        | 	pivot_pose = pose_trans(p_center, hinge_offset)
        | 	pose_rel = pose_trans(pose_inv(pivot_pose), p_center)
        | 	angle_mid = (angle/2.0)*3.1416/180
        | 	angle_end = angle*3.1416/180
        | 	tilt_mid = p[0,0,0, -angle_mid, 0, 0]
        | 	tilt_end = p[0,0,0, -angle_end, 0, 0]
        | 	pose_rel_mid = pose_trans(tilt_mid, pose_rel)
        | 	pose_rel_end = pose_trans(tilt_end, pose_rel)
        | 	via_pose = pose_trans(pivot_pose, pose_rel_mid)
        | 	end_pose = pose_trans(pivot_pose, pose_rel_end)
        | 	movec(via_pose, end_pose, a=0.05, v=0.01, r=0.001)
        | 	p_center = get_actual_tcp_pose()
        | end
        | 
        | def deg2rad(d):
        | 	return d*3.141592/180
        | end
        | 
        | def map_tilt_to_ry_deg(container_deg):
        | 
        | 	if (Flowability == "Easy" or Flowability == "Medium"):
        | 		if ( level>=10.0):
        | 			ry_min = 10.0
        | 			ry_max = 75.0
        | 		elif (level<10.00 and level >1.00):
        | 			ry_min = 16.0
        | 			ry_max = 65.0
        | 		else:
        | 			ry_min=17.0
        | 			ry_max=75.0
        | 		end
        | 	else:
        | 		if ( level>=10.0):
        | 			ry_min = 0.0
        | 			ry_max = 65.0
        | 		elif (level<10.00 and level >1.00):
        | 			ry_min = 10.0
        | 			ry_max = 45.0
        | 		else:
        | 			ry_min=0.0
        | 			ry_max=50.0
        | 		end
        | 
        | 	end
        | 
        | 	local span_count = angle_max -angle_min
        | 	local span_ry = ry_max - ry_min
        | 
        | 	local t = (container_deg -angle_min)/span_count
        | 	local ry_deg = ry_max - t*span_ry
        | 
        | 	return clamp(ry_deg, ry_min, ry_max)
        | 
        | end
        | 
        | def caluclate_corrections(level):
        | 	z_high = 0.01
        | 	z_low = -0.08
        | 	y_high = -0.01
        | 	y_low = -0.015
        | 
        | 	scale = (level - 10.0) / (100.0-10.0)
        | 
        | 	global correction_z = z_low + scale*(z_high - z_low)
        | 	global correction_y = y_low + scale*(y_high -y_low)
        | 
        | end
        | 
        | def scoop_powder(p_center):
        | 	#lift_offset = p[0, 0, 0.05, 0, 0, 0]
        | 	vibration_voltage = 0.4
        | 	vibration_time = 3.0
        | 	diameter = 0.07
        | 	global scoop_radius_default = 0.0
        | 	#p_center = center_pose_t
        | 
        | 
        | 	if (level >=70.00):
        | 		approach_offset = p[0.008,0,0.22,0,0,0]
        | 		lift_offset = p[0, 0, 0.05, 0, 0, 0]
        | 		caluclate_corrections(level)
        | 	elif (level >=10.00 and level <70):
        | 		approach_offset = p[0.008,0,0.22,0,0,0]
        | 		lift_offset = p[0, 0, 0.15, 0, 0, 0]
        | 		caluclate_corrections(level)
        | 	elif (level<10.00 and level >= 1.00):
        | 		approach_offset = p[0.01,0,0.22,0,0,0]
        | 		correction_z = -0.08
        | 		correction_y = -0.01
        | 		lift_offset = p[0, 0, 0.14, 0, 0, 0]
        | 	else:
        | 		approach_offset = p[0.008,0,0.22,0,0,0]
        | 		correction_z = -0.08
        | 		correction_y = -0.01
        | 		lift_offset = p[0, 0, 0.14, 0, 0, 0]
        |  	end
        | 
        | 	if (spatula == "spatula_L"):
        | 		global spatula_depth = 0.015
        | 	elif (spatula == "spatula_M"):
        | 		global spatula_depth = 0.01
        | 	elif (spatula == "spatula_S"):
        | 		global spatula_depth = 0.008
        | 	elif (spatula == "spatula_flat_M"):
        | 		global spatula_depth = 0.001
        | 	elif (spatula == "spatula_flat_S"):
        | 		global spatula_depth = 0.005
        | 	end
        | 
        | 	scoop_radius_default = diameter/2 - spatula_depth
        | 	scoop_entry_pose = pose_trans(p_center, approach_offset)
        | 	movel(scoop_entry_pose, a=0.1, v=0.25)
        | 
        | 	scoop_start_rel = p[scoop_radius_default, 0, scoop_depth, 0, 0, 0]
        | 
        | 	rot_mid = p[0, 0, 0, 0, 0, 0.785]
        | 	rot_end = p[0, 0, 0, 0, 0, 1.5708]
        | 
        | 	scoop_via_rel = pose_trans(rot_mid, scoop_start_rel)
        | 	scoop_end_rel = pose_trans(rot_end, scoop_start_rel)
        | 
        | 	scoop_start_pose = pose_trans(p_center, scoop_start_rel)
        | 	scoop_via_pose = pose_trans(p_center, scoop_via_rel)
        | 	scoop_end_pose = pose_trans(p_center, scoop_end_rel)
        | 
        | 	movel(scoop_start_pose, a=0.5, v=0.3)
        | 	#movel(p_center, a=0.5, v=1.0)
        | 	#sleep(5.0)
        | 
        | 	if (level<90.0):
        | 		Rotate()
        | 	end
        | 
        | 	#movec(scoop_via_pose, scoop_end_pose, a=0.03, v=0.05)
        | 	movec(scoop_via_pose, scoop_end_pose, a=0.03, v=0.02)
        | 	#movel(pose_trans(get_actual_tcp_pose(), p[0,0,0,0,0,deg2rad(90.0)]), a=0.03, v=0.05)
        | 	sleep(1.0)
        | 	local ry_deg = map_tilt_to_ry_deg(angle_deg)
        | 	local ry = deg2rad(ry_deg)
        | 	local end_rel = pose_trans(pose_inv(p_center), scoop_end_pose)
        | 	local end_rel_tilted = pose_trans(end_rel, p[0, 0, 0, 0, ry, 0])
        | 	global tilted_pose_in_base = pose_trans(p_center, p[0,correction_y,correction_z,end_rel_tilted[3],end_rel_tilted[4], end_rel_tilted[5]])
        | 	global tilted_pose_in_base = pose_trans(tilted_pose_in_base, p[0, 0, spatula_len, 0, 0, 0])
        | 
        | 	if (Flowability == "Hard"):
        | 		tilt_send((angle_deg+5))
        | 	end
        | 	movel(tilted_pose_in_base, a=0.03, v=0.1)
        | 
        | 	if (Flowability == "Hard"):
        | 		tilt_send((angle_deg-5))
        | 	end
        | 
        | 	if (spatula=="spatula_flat_S" or spatula=="spatula_S"):
        | 		vibration_3()
        | 	else:
        | 		set_analog_out(0, vibration_voltage)
        | 	end
        | 	if (Flowability == "Easy"):
        | 		local n=1.4
        | 	else:
        | 		local n=1.5
        | 	end
        | 	local ry_level = deg2rad(ry_deg/n)
        | 	local end_rel_tilted_level = pose_trans(end_rel, p[0, 0, 0, 0, ry_level, 0])
        | 	local level_tilted_pose_in_base = pose_trans(p_center, p[0,correction_y,correction_z,end_rel_tilted_level[3],end_rel_tilted_level[4], end_rel_tilted_level[5]])
        | 	local level_tilted_pose_in_base = pose_trans(level_tilted_pose_in_base, p[0, 0, spatula_len, 0, 0, 0])
        | 
        | 	movel(level_tilted_pose_in_base, a=0.03, v=0.1)
        | 	#if (level>70.0):
        | 		#sleep(1.0)
        | 	#end
        | 	sleep(1.0)
        | 	#sleep(vibration_time)
        | 
        | 	movel(tilted_pose_in_base, a=0.03, v=0.1)
        | 	set_analog_out(0, 0.0)
        | 
        | 	tilt_pose_rel = pose_trans(pose_inv(p_center), tilted_pose_in_base)
        | 
        | 	lifted_pose_rel = pose_trans(lift_offset, tilt_pose_rel)
        | 
        | 	global lifted_pose = pose_trans(p_center, lifted_pose_rel)
        | 	movel(lifted_pose, a=0.03, v=0.1)
        | 	CCW_Rotate()
        | end
        | 
        | 
        | def center_pose():
        | 	trans_rel = p[0.0, 0.05, 0.0, 0, 0, 0]
        | 
        | 	p_translated = pose_trans(place_pose, trans_rel)
        | 	cx = p_translated[0]
        | 	cy = p_translated[1]
        | 	cz = p_translated[2]
        | 
        | 	global p_center_vertical = p[cx,cy,cz, 0, 0, 4.09]
        | 
        | 	#movej(p_center_vertical, a =0.3, v =0.3)
        | 	#sleep(3.0)
        | 	return p_center_vertical
        | end
        | 
        | def updated_center_pose(p_center_vertical, angle_deg):
        | 	hinge_pose = pose_trans(p_center_vertical, p[0,0,-0.2,0,0,0])
        | 	local_rel = pose_trans(pose_inv(hinge_pose), p_center_vertical)
        | 
        | 	rot_tilt = p[0,0,0, -deg2rad(angle_deg),0,0]
        | 	local_rel_tilted = pose_trans(rot_tilt, local_rel)
        | 
        | 	global p_center = pose_trans(hinge_pose, local_rel_tilted)
        | 	return p_center
        | end
        | 
        | def tilt_send(angle):
        | 	socket_open("192.168.12.101", 80)
        | 	angle = 92.0 - angle
        | 	socket_send_string("Tilt,"+to_str(angle)+",0")
        | 	sync()
        | 	sleep(0.5)
        | 	socket_close()
        | end
        | 
        | def Motors_off():
        | 	socket_open("192.168.12.101", 80)
        | 	socket_send_string("Off,0,0")
        | 	sync()
        | 	sleep(0.5)
        | 	socket_close()
        | end
        | 
        | def Rotate():
        | 	socket_open("192.168.12.101", 80)
        | 	socket_send_string("FullRotation, 1, 2000")
        | 	sync()
        | 	sleep(0.5)
        | 	socket_close()
        | end
        | 
        | 
        | def CCW_Rotate():
        | 	socket_open("192.168.12.101", 80)
        | 	socket_send_string("FullRotation, -1, 2000")
        | 	sync()
        | 	sleep(0.5)
        | 	socket_close()
        | end
        | def tilt_to_home():
        | 	socket_open("192.168.12.101", 80)
        | 	socket_send_string("Home,0,0")
        | 	sync()
        | 	sleep(0.5)
        | 	socket_close()
        | end
    Script file /programs/04 Scripts/Weight_scale_socket.script
      | def get_weight():
      | 	socket_open("192.168.12.111", 3002)
      | 	sleep(0.2)
      | 	textmsg("socket opened successfully!")
      | 	socket_send_string("GET_WEIGHT")
      | 	sync()
      | 	sleep(0.5)
      | 	receiveFromServ = socket_read_ascii_float(6)
      | 	while (receiveFromServ[0] <1):
      | 		sleep(0.5)
      | 		receiveFromServ = socket_read_ascii_float(1)
      | 		textmsg("retrying read:", receiveFromServ)
      | 	end
      | 	textmsg("Received weight:", receiveFromServ[1])
      | 	socket_close()
      | 	sleep(0.2)
      | 	return receiveFromServ[1]
      | end
      | 
      | def tare_scale():
      | 	socket_open("192.168.12.111", 3002)
      | 	socket_send_string("TARE")
      | 	sleep(0.5)
      | 	socket_close()
      | end
      | 
      | def zero_scale():
      | 	socket_open("192.168.12.111", 3002)
      | 	socket_send_string("ZERO")
      | 	sleep(0.5)
      | 	socket_close()
      | end
      | 
      | def log_weight():
      | 	socket_open("192.168.12.111", 3002)
      | 	socket_send_string("LOG_WEIGHT")
      | 	sleep(0.5)
      | 	socket_close()
      | end
      | 
      | def send_target_info():
      | 	socket_open("192.168.12.111", 3002)
      | 	socket_send_string("SET_TARGET:" + to_str(target_weight))
      | 	sleep(0.2)
      | 	socket_close()
      | end
      | def send_powder_info():
      | 	socket_open("192.168.12.111", 3002)
      | 	socket_send_string("SET_POWDER:" + Pow_name)
      | 	sleep(0.2)
      | 	socket_close()
      | end
      | def send_spatula_info():
      | 	socket_open("192.168.12.111", 3002)
      | 	socket_send_string("SET_SPATULA:" + spatula)
      | 	sleep(0.2)
      | 	socket_close()
      | end
      | 
      | def send_level_info():
      | 	socket_open("192.168.12.111", 3002)
      | 	socket_send_string("SET_LEVEL:" + to_str(level))
      | 	sleep(0.2)
      | 	socket_close()
      | end
      | def Dosing_done():
      | 	socket_open("192.168.12.111", 3002)
      | 	socket_send_string("DOSING_DONE")
      | 	sleep(0.2)
      | 	socket_close()
      | end
      | 
      | def send_dosing_time(Dosed_time):
      | 	socket_open("192.168.12.111", 3002)
      | 	socket_send_string("DOSED_TIME:" + to_str(Dosed_time))
      | 	sleep(0.2)
      | 	socket_close()
      | end
    Script file /programs/04 Scripts/Calibration.script
      | # ------------------------------------------------------------
      | # Theoretical W_FULL from Cylinder Volume + Density
      | # (Eliminates manual W_FULL; keeps W_EMPTY + W_now for level)
      | # ------------------------------------------------------------
      | # -------------------------
      | # 1) Define container geometry (cylindrical inner dimensions)
      | # -------------------------
      | # Use mm for readability; we convert internally.
      | global D_INNER_MM   = 66.0     # inner diameter of container (mm)
      | global H_FILL_MM    = 125.0    # usable fill height up to "full" (mm)
      | 
      | # -------------------------
      | # 2) Define powder density
      | # -------------------------
      | # Density is directly set for now (as per your requirement).
      | # Use g/mL (common lab bulk density style).
      | #global RHO_G_PER_ML = 0.40     # example: 0.55 g/mL (replace per powder)
      | 
      | # ------------------------------------------------------------
      | # Spatula volumes (manufacturer specified)
      | # ------------------------------------------------------------
      | 
      | # Large spatula
      | global SPATULA_L_VOL_ML = 5.0        # 1 teaspoon = 5 mL
      | 
      | # Medium spatula
      | global SPATULA_M_VOL_ML = 1.25       # 1/4 teaspoon = 1.25 mL
      | 
      | # Small spatula
      | global SPATULA_S_VOL_ML = 0.15625    # 1/32 teaspoon = 0.15625 mL
      | 
      | global SPATULA_FLAT_M_VOL_ML  = 2.2
      | global SPATULA_FLAT_S_VOL_ML  = 1.2   #based on caluclations using rho = m/V
      | 
      | # -------------------------
      | # 4) Utility functions
      | # -------------------------
      | 
      | 
      | def cyl_volume_mL(d_mm, h_mm):
      |   # Converts mm -> m, computes cylinder volume in m^3, converts to mL
      |   # V = π * r^2 * h
      |   local d_m  = d_mm / 1000.0
      |   local h_m  = h_mm / 1000.0
      |   local r_m  = d_m / 2.0
      |   local v_m3 = 3.141592653589793 * r_m * r_m * h_m
      |   global v_mL = v_m3 * 1000000.0     # 1 m^3 = 1,000,000 mL
      |   return v_mL
      | end
      | 
      | def compute_W_full_theoretical():
      |   V_mL = cyl_volume_mL(D_INNER_MM, H_FILL_MM)
      |   local M_powder_g = density * V_mL
      |   global W_FULL = W_EMPTY + M_powder_g
      |   return W_FULL
      | end
      | 
      | 
      | # ------------------------------------------------------------
      | # Function: Theoretical scoop weight from volume
      | # ------------------------------------------------------------
      | def scoop_weight_from_volume(vol_mL, density):
      |   return vol_mL * density
      | end
      | 
      | # ------------------------------------------------------------
      | # Function: Get scoop weight based on spatula type
      | # ------------------------------------------------------------
      | def get_scoop_weight(spatula):
      |   local vol = 0.0
      | 
      |   if (spatula == "spatula_L"):
      |     vol = SPATULA_L_VOL_ML
      |   elif (spatula == "spatula_M"):
      |     vol = SPATULA_M_VOL_ML
      |   elif (spatula == "spatula_S"):
      |     vol = SPATULA_S_VOL_ML
      |   elif (spatula == "spatula_flat_M"):
      |     return SPATULA_FLAT_M_VOL_ML
      |   elif (spatula == "spatula_flat_S"):
      |     return SPATULA_FLAT_S_VOL_ML
      |   else:
      |     textmsg("Unknown spatula type")
      |     return 0.0
      |   end
      | 
      |   global target_g =  scoop_weight_from_volume(vol, density)
      |   return target_g
      | end
  Folder BeforeStarts [hidden by the author, left out]
  Folder powder dispensing variable init
    Start_thread := False
    vib_thread := False
    kp := 0.001
    ki := 0.00006
    kd := 0.015
    dt := 0.03
    Integral_error := 0
    current_error := 0
    previous_error := 0
    tilt_increment := 0
    tilt_angle := 0
    diff := 0
    current_pose := get_actual_tcp_pose()
    Relative_trans := p[0, 0, -0.035, 0, 0, 0]
    ContA_plc_offst := p[-0.00205, 0.02547, 0.03730, -0.03, -2.183, 6.165]
    PowA_50_offset := p[0.21808, -0.19943, 0.06584, 0, 0, 0]
    SuppressedNode
      Script: scooping_init()
    Script: tilt_init_reference()
    switch_spat_M := True
    switch_spat_S := True
    switch_spat_F_M := True
    switch_spat_F_S := True
    last_scale := 0
    W_EMPTY := 51.3
    w_dosed_total := 0
Robot Program (runOnlyOnce=false)
  Folder MAIN
    Script: command_manager(external_control="uGO", cond_suspend=(ITM_Manipulated and AMR_AtTarget and AMR_Charging and AMR_Battery<40), cond_unsuspend=(AMR_Battery≟60))
    Script: log_state(STATE_Info)
    Switch expression=STATE
      Case (caseValue=1)
        Folder Stopping
          STATE_Info := "Stopping"
          Script: end_freedrive_mode()
          Set NoAction tcp=TCP
          PSE_T := get_tool_free_pose(dir=[0,0,0.150], move_in_base_frame=True)
          If is_reachable(Base, [PSE_T])
            MoveL speed 150 mm/s, acceleration 1200 mm/s^2 (useActiveTCP=true optimoveEnabled=false optiMoveSpeed=0.3 optiMoveAcceleration=0.09) feature=Base
              Waypoint Variable (Variable): variable=PSE_T
          Script: do_transition(keep_rxry=OBJ_Picked, r=0)
          SuppressedNode
            Folder Decapper
              Set DigitalOutput pin=digital_out[4]; digitalValue=0
              Set DigitalOutput pin=BarcodeTrigger; digitalValue=0
              Set DigitalOutput pin=digital_out[3]; digitalValue=0
              Set DigitalOutput pin=digital_out[2]; digitalValue=0
              Set DigitalOutput pin=digital_out[5]; digitalValue=0
          SuppressedNode
            Folder Centrifuge [hidden by the author, left out]
          Call Sub_AMR_MiR_V3
          If stopping() and AMR_Done
            STATE := 2
            Script: ugo_update_outputs()
      Case (caseValue=2)
        Folder Stopped
          STATE_Info := "Stopped"
          Call Sub_AMR_MiR_V3
          If CMD_Reset  or PB_Start
            STATE := 3
            Script: ugo_update_outputs()
      Case (caseValue=3)
        Folder  Resetting [hidden by the author, left out]
      Case (caseValue=4)
        Folder Idle [hidden by the author, left out]
      Case (caseValue=5)
        Folder Starting
          STATE_Info := "Starting"
          'ADD COMMANDS WHAT TO START WITH'
          Call Sub_AMR_MiR_V3
          Folder get ugo data
            Folder Assign Tasks
              Script: TASK.ID = ugo_get_task()
              If TASK.ID≟1
                Task_info := "Charge"
                Folder Parameters
                  AMR_PosTarget := 1
              ElseIf TASK.ID≟9
                'Pick Sarstedt Rack from Variable source'
                Task_info := "Navigate to Target"
                Folder Parameters
                  AMR_PosTarget := UGO.read_input("00","ITM_ID")
              ElseIf TASK.ID≟49
                Task_info := "Pick Containers"
                Folder Parameters
                  ITM_ID := 1
                  OBJ_Type := 6
                  JIG := 15
                  AMR_PosTarget := 3
              ElseIf TASK.ID≟50
                Task_info := "Decap Containers"
                Folder Parameters
                  ITM_ID := 1
                  OBJ_Type := 6
                  JIG := 16
                  AMR_PosTarget := 5
              ElseIf TASK.ID≟51
                Task_info := "Detect Spatula and transfer powder"
                Folder Parameters
                  ITM_ID := 1
                  target_weight := (UGO.read_input("00","Target_weight"))/1000
                  OBJ_Type := 8
                  JIG := 16
                  AMR_PosTarget := 5
              ElseIf TASK.ID≟52
                Task_info := "Pick Powder"
                Folder Parameters
                  ITM_ID := 1
                  OBJ_Type := 6
                  JIG := 15
                  AMR_PosTarget := 3
              ElseIf TASK.ID≟53
                Task_info := "Decap Powder"
                Folder Parameters
                  ITM_ID := 1
                  OBJ_Type := 6
                  JIG := 1
                  AMR_PosTarget := 5
              ElseIf TASK.ID≟54
                Task_info := "Empty and swap Powder container"
                SuppressedNode
                  Folder Parameters
                    ITM_ID := 1
                    target_weight := (UGO.read_input("00","Target_weight"))/1000
                    W_now := (UGO.read_input("00","Container_weight"))/1000
                    Pow_name := (UGO.read_input("00","Powder_name"))
                    OBJ_Type := 6
                    JIG := 17
                    AMR_PosTarget := 5
                Folder Parameters
                  ITM_ID := 1
                  SuppressedNode
                    target_weight := (UGO.read_input("00","target_weight"))/1000
                  W_now := (UGO.read_input("00","Container_weight"))/1000
                  Pow_name := (UGO.read_input("00","Powder_name"))
                  Script: scooping_init()
                  target_weight := W_now-W_EMPTY-(0.002*W_FULL)
                  OBJ_Type := 6
                  JIG := 17
                  AMR_PosTarget := 5
              ElseIf TASK.ID≟55
                Task_info := "Place Powder"
                Folder Parameters
                  ITM_ID := 1
                  OBJ_Type := 6
                  JIG := 21
                  AMR_PosTarget := 5
              ElseIf TASK.ID≟56
                Task_info := "Dose Powder"
                Folder Parameters
                  ITM_ID := 1
                  target_weight := (UGO.read_input("00","Target_weight"))/1000
                  W_now := (UGO.read_input("00","Container_weight"))/1000
                  SuppressedNode
                    W_now := 135
                  Pow_name := (UGO.read_input("00","Powder_name"))
                  OBJ_Type := 6
                  JIG := 17
                  AMR_PosTarget := 5
              ElseIf TASK.ID≟57
                Task_info := "Recipe Powder dosing"
                Folder Parameters
                  ITM_ID := 1
                  Pow_A := (UGO.read_input("00","PowderA"))
                  Pow_B := (UGO.read_input("00","PowderB"))
                  Pow_C := (UGO.read_input("00","PowderC"))
                  Total_weight := (UGO.read_input("00","Total_weight"))/1000
                  Pow_A_percent := (UGO.read_input("00","PowderA_percentage"))/100
                  Pow_B_percent := (UGO.read_input("00","PowderB_percentage"))/100
                  Pow_C_percent := (UGO.read_input("00","PowderC_percentage"))/100
                  OBJ_Type := 6
                  JIG := 17
                  AMR_PosTarget := 5
              ElseIf TASK.ID≟58
                Task_info := "Pick Powder containers"
                Folder Parameters
                  ITM_ID := 1
                  OBJ_Type := 6
                  JIG := 15
                  AMR_PosTarget := 3
              ElseIf TASK.ID≟59
                Task_info := "Calibration for new powder"
                Folder Parameters
                  ITM_ID := 1
                  Pow_name := (UGO.read_input("00","Pow_name"))
                  W_now := (UGO.read_input("00","Container_weight"))/1000
                  density := (UGO.read_input("00", "Density"))
                  Flowability := (UGO.read_input("00", "Flowability"))
                  spatula := (UGO.read_input("00","Spatula"))
                  OBJ_Type := 6
                  JIG := 17
                  AMR_PosTarget := 5
              Else 
                Script: set_error(ERROR_WRONG_ORDER)
          Folder test ugo
            Wait Sleep waitTime=0.2
            Script: ugo_update_outputs()
          If starting() and AMR_Done
            Script: log_message(Task_info, "New Task: ")
            Script: log_message(to_str(TASK.ID), "Task_ID: ")
            Script: do_transition(keep_rxry=OBJ_Picked)
            STATE := 6
            Script: ugo_update_outputs()
      Case (caseValue=6)
        Folder Execute
          STATE_Info := "Execute"
          If not CMD_Hold and not CMD_Suspend (checkContinuously=true)
            Switch expression=PROCESS_Step
              Case (caseValue=0)
                PROCESS_Info := "process control"
                Script: log_process(PROCESS_Info)
                Folder process control [hidden by the author, left out]
              Case (caseValue=1)
                Folder navigate
                  'MOVING THE uML'
                  PROCESS_Info := "move to target"
                  Script: log_process(PROCESS_Info)
                  If TASK.ID≟1
                    Action := 51
                  Else 
                    Action := 52
                  Call Sub_AMR_MiR_V3
                  If AMR_Done
                    PROCESS_Step := 0
              Case (caseValue=2)
                Folder prepare
                  'THINGS THAT HAVE TO BE DONE ONCE IN A SEQUENCE,WORKFLOW'
                  PROCESS_Info := "prepare for work"
                  Script: log_process(PROCESS_Info)
                  If TASK.WORK.ITM_ID_Src>1
                    ITM_ID := TASK.WORK.ITM_ID_Src
                  ElseIf TASK.WORK.ITM_ID_Tgt>1
                    ITM_ID := TASK.WORK.ITM_ID_Tgt
                  If not ARM_Referenced and (ITM_ID≠0)
                    STP := 1
                  ElseIf ARM_Referenced or (ITM_ID≟0)
                    STP := 2
                  Switch expression=STP
                    Case (caseValue=1)
                      Folder reference
                        STP_Info := "reference at target position"
                        Script: log_step(STP_Info)
                        If ITM_ID≟1
                          CAM_Done := True
                        Else 
                          Action := 131
                          Call Sub_Vision_V18
                          SuppressedNode
                            CAM_Done := True
                        If CAM_Done and  not ERROR.FLAG
                          Script: log_step("ARM referenced")
                          ARM_Referenced := True
                    Case (caseValue=2)
                      Folder manipulate [hidden by the author, left out]
                  ITM_Prepared := (ITM_Manipulated or  not found_in_list(ITM_ID, ITM_ID_List)) and (ARM_Referenced or ITM_ID≟0) and  not WRK_Done
                  STP := 0
                  STP_Info := ""
                  PROCESS_Step := 0
              Case (caseValue=3)
                Folder work
                  'ADD EVERY MACHINE, OBJECT, STATION TO WORK ON'
                  Switch expression=ITM_ID
                    Case (caseValue=1)
                      Folder uLM
                        If TASK.ID≟12
                          Folder fill racks
                            Action := 151
                            Call Sub_Vision_V18
                            If not ERROR.FLAG
                              Folder Actions for the task
                                Action := 1
                                JIG := 2
                                JIG_Slot := CAM_Result[0]
                                OBJ_Nbr := CAM_Result[0]
                                OBJ_Type := 2
                                Call Sub_Action_V4
                                If OBJ_Picked
                                  Script: CAM_Result.remove(0)
                                  PRC_TubCounter := PRC_TubCounter+1
                                  If PRC_TubCounter%4≟0
                                    JIG_Slot := 4
                                  Else 
                                    JIG_Slot := PRC_TubCounter%4
                                  OBJ_Nbr := ceil(PRC_TubCounter/4)
                                  Action := 2
                                  JIG := 4
                                  Call Sub_Action_V4
                                  Action := 151
                                  Call Sub_Vision_V18
                            If (CAM_Captures≥CAM_PRM_Retries) or (PRC_TubCounter≥32)
                              PROCESS_Step := 0
                              WRK_Done := True
                        ElseIf TASK.ID≟49
                          Folder Pick Powder container
                            Action := 131
                            Call Sub_Vision_V18
                            Action := 35
                            Call Sub_Action_V4
                            PROCESS_Step := 0
                            WRK_Done := True
                        ElseIf TASK.ID≟50
                          Folder Decap containers
                            Action := 36
                            Call Sub_Action_V4
                            PROCESS_Step := 0
                            WRK_Done := True
                        ElseIf TASK.ID≟51
                          Folder Detect Spatula and transfer powder
                            Action := 131
                            Call Sub_Vision_V18
                            Action := 37
                            Call Sub_Action_V4
                            PROCESS_Step := 0
                            WRK_Done := True
                        ElseIf TASK.ID≟52
                          Folder Pick Powder container
                            Action := 131
                            Call Sub_Vision_V18
                            Action := 39
                            Call Sub_Action_V4
                            PROCESS_Step := 0
                            WRK_Done := True
                        ElseIf TASK.ID≟53
                          Folder Decap containerA
                            Action := 40
                            Call Sub_Action_V4
                            PROCESS_Step := 0
                            WRK_Done := True
                        ElseIf TASK.ID≟55
                          Folder Place Powder
                            Action := 131
                            Call Sub_Vision_V18
                            Action := 41
                            Call Sub_Action_V4
                            PROCESS_Step := 0
                            WRK_Done := True
                        ElseIf TASK.ID≟54
                          Folder Empty and swap container
                            Action := 131
                            Call Sub_Vision_V18
                            Action := 42
                            Call Sub_Action_V4
                            PROCESS_Step := 0
                            WRK_Done := True
                        ElseIf TASK.ID≟56
                          Folder Dispense Powder
                            Action := 131
                            Call Sub_Vision_V18
                            Action := 43
                            Call Sub_Action_V4
                            PROCESS_Step := 0
                            WRK_Done := True
                        ElseIf TASK.ID≟57
                          Folder Recipe Dosing
                            QR_Action := 1
                            Action := 48
                            Call Sub_Action_V4
                            Script: recipe_init(Pow_A, Pow_B, Pow_C, Total_weight, Pow_A_percent, Pow_B_percent, Pow_C_percent)
                            Loop While (checkContinuously=false) expression=recipe_next()≟ True
                              Action := 44
                              Call Sub_Action_V4
                              JIG := 21
                              Action := 131
                              Call Sub_Vision_V18
                              Action := 45
                              Call Sub_Action_V4
                              Script: dosing_start()
                              JIG := 17
                              Action := 131
                              Call Sub_Vision_V18
                              Action := 46
                              Call Sub_Action_V4
                              Script: dosing_end()
                            PROCESS_Step := 0
                            WRK_Done := True
                        ElseIf TASK.ID≟58
                          Folder Pick Powder containers
                            Num_cont_picked := 0
                            powder_position := "Position1"
                            Loop While (checkContinuously=false) expression=Num_cont_picked<3
                              Action := 131
                              Call Sub_Vision_V18
                              Action := 47
                              Call Sub_Action_V4
                            PROCESS_Step := 0
                            WRK_Done := True
                        ElseIf TASK.ID≟59
                          Folder Calibration
                            SuppressedNode
                              QR_Action := 2
                            SuppressedNode
                              Action := 48
                            SuppressedNode
                              Call Sub_Action_V4
                            Action := 49
                            Call Sub_Action_V4
                            PROCESS_Step := 0
                            WRK_Done := True
                    Case (caseValue=2)
                      SuppressedNode
                        Folder Centrfiuge
                          SuppressedNode
                            Script: cent_error_check()
                          OBJ_Type := 1
                          If not ERROR.FLAG
                            'load racks'
                            If TASK.ID≟14
                              Loop While (checkContinuously=false) expression=(PRC_RackCounter<4) and  not CMD_Stop and  not ERROR.FLAG
                                ITM_ID := TASK.WORK.ITM_ID_Src
                                JIG := 4
                                JIG_Slot := PRC_RackCounter+1
                                Action := 1
                                CallSubProgram
                                If OBJ_Picked and  not ERROR.FLAG
                                  ITM_ID := TASK.WORK.ITM_ID_Tgt
                                  Script: execute_cent_action(ACTION_ROTATE, JIG_Slot)
                                  Action := 7
                                  CallSubProgram
                                  PRC_RackCounter := PRC_RackCounter + 1
                              If not ERROR.FLAG
                                WRK_Done := True
                                PROCESS_Step := 0
                            'unload racks'
                            If TASK.ID≟15
                              If CNT_State_Actual≟2 or CNT_State_Actual≟3
                                Loop While (checkContinuously=false) expression=(PRC_RackCounter<4) and  not CMD_Stop and  not ERROR.FLAG
                                  ITM_ID := TASK.WORK.ITM_ID_Src
                                  JIG_Slot := PRC_RackCounter + 1
                                  Script: execute_cent_action(ACTION_ROTATE, JIG_Slot)
                                  Script: execute_cent_action(ACTION_INSPECT, JIG_Slot)
                                  Action := 8
                                  CallSubProgram
                                  If OBJ_Picked and  not ERROR.FLAG
                                    ITM_ID := TASK.WORK.ITM_ID_Tgt
                                    JIG := 4
                                    JIG_Slot := PRC_RackCounter + 1
                                    Action := 2
                                    CallSubProgram
                                    PRC_RackCounter := PRC_RackCounter+1
                                If not ERROR.FLAG
                                  WRK_Done := True
                                  PROCESS_Step := 0
                    Case (caseValue=5)
                      SuppressedNode
                        Folder SarstedtTable
                          Action := 131
                          CallSubProgram
                          Action := 1
                          CallSubProgram
                          PROCESS_Step := 0
                          WRK_Done := True
                    Case (caseValue=20)
                      SuppressedNode
                        Folder Biorad rack
                          'load racks'
                          If Task_ID≟16
                            SuppressedNode
                              PRC_RackCounter := 0
                            Loop While (checkContinuously=false) expression=(PRC_RackCounter<PRC_RackNumber) and  not CMD_Stop
                              JIG_Slot := PRC_RackCounter
                              Action := 1
                              PRC_Target := 0
                              CallSubProgram
                              If OBJ_Picked
                                Action := 2
                                PRC_Target := 1
                                CallSubProgram
                                Action := 7
                                PRC_Target := 1
                                CallSubProgram
                                PRC_RackCounter := PRC_RackCounter+1
                            WRK_Done := True
                            PROCESS_Step := 0
                          'unload racks'
                          SuppressedNode
                            If Task_ID≟17
                              SuppressedNode
                                PRC_RackCounter := 0
                              Loop While (checkContinuously=false) expression=(PRC_RackCounter<PRC_RackNumber) and  not CMD_Stop
                                JIG_Slot := PRC_RackCounter
                                Action := 8
                                PRC_Target := 1
                                Script: textmsg("Callactionunload=",Action)
                                CallSubProgram
                                Action := 1
                                PRC_Target := 1
                                Script: textmsg("Callactionpick=",Action)
                                CallSubProgram
                                If OBJ_Picked
                                  Action := 2
                                  PRC_Target := 0
                                  Script: textmsg("Callactionplace=",Action)
                                  CallSubProgram
                                  PRC_RackCounter := PRC_RackCounter+1
                              WRK_Done := True
                              PROCESS_Step := 0
                          If Task_ID≟17
                            PRC_RackCounter := 0
                            Loop While (checkContinuously=false) expression=(PRC_RackCounter<PRC_RackNumber) and  not CMD_Stop
                              Wait Condition expression=SensorData[PRC_RackCounter]≟1
                              JIG_Slot := PRC_RackCounter
                              Action := 8
                              PRC_Target := 1
                              Script: textmsg("Callactionunload=",Action)
                              CallSubProgram
                              Action := 1
                              PRC_Target := 1
                              Script: textmsg("Callactionpick=",Action)
                              CallSubProgram
                              If OBJ_Picked
                                Action := 2
                                PRC_Target := 0
                                Script: textmsg("Callactionplace=",Action)
                                CallSubProgram
                                PRC_RackCounter := PRC_RackCounter+1
                            WRK_Done := True
                            PROCESS_Step := 0
                    Case (caseValue=43)
                      SuppressedNode
                        Folder Pick the rack
                          Action := 131
                          CallSubProgram
                          Action := 1
                          CallSubProgram
                          PROCESS_Step := 0
                          WRK_Done := True
                    Case (caseValue=2147483647)
                      WRK_Done := True
                      PROCESS_Step := 0
          If CMD_Hold
            STATE := 9
            Script: ugo_update_outputs()
          ElseIf CMD_Suspend
            STATE := 12
            Script: ugo_update_outputs()
      Case (caseValue=7)
        Folder Completing [hidden by the author, left out]
      Case (caseValue=8)
        Folder Complete [hidden by the author, left out]
      Case (caseValue=9)
        Folder Holding [hidden by the author, left out]
      Case (caseValue=10)
        Folder Held [hidden by the author, left out]
      Case (caseValue=11)
        Folder Unholding [hidden by the author, left out]
      Case (caseValue=12)
        Folder Suspending [hidden by the author, left out]
      Case (caseValue=13)
        Folder Suspended [hidden by the author, left out]
      Case (caseValue=14)
        Folder Unsuspending [hidden by the author, left out]
      Case (caseValue=15)
        Folder Aborting [hidden by the author, left out]
      Case (caseValue=16)
        Folder Aborted [hidden by the author, left out]
      Case (caseValue=17)
        Folder Clearing [hidden by the author, left out]
    Script: log_state(STATE_Info)
    Script: log_warning(WARNING.MSG)
    Script: log_error(ERROR.MSG)
    Folder Times [hidden by the author, left out]
    SuppressedNode
      Script: sync()
    Wait Sleep waitTime=0.1
Thread Thread_1 (runOnlyOnce=false)
  If Start_thread≟ True
    weight_value := get_weight()
    Wait Sleep waitTime=0.1
    Script: sync()
  Script: sync()
Thread Thread_2 (runOnlyOnce=false)
  Loop While (checkContinuously=true) expression=vib_thread≟ True
    diff := target_weight-weight_value
    If diff>0.02 and spatula≠"spatula_flat_S" (checkContinuously=true)
      SuppressedNode
        Script: vibration_1()
      Set AnalogOutput pin=analog_out[0]; analogValue=4
    ElseIf diff>0.02 and spatula≟"spatula_flat_S"
      Script: vibration_3()
    ElseIf diff≤0.03 (checkContinuously=true)
      Script: vibration_2()
    SuppressedNode
      ElseIf diff≥0.01 and diff<0.05
        Script: vibration_3()
    SuppressedNode
      ElseIf diff>0 and diff<0.01
        Script: vibration_4()
    Else 
      Set AnalogOutput pin=analog_out[0]; analogValue=0
  Script: sync()
SubProgram -> Sub_Vision_V18
SubProgram  [hidden by the author, left out]
SubProgram -> Sub_Action_V4
SubProgram Sub_AMR_MiR_V3 [hidden by the author, left out]
SubProgram Sub_Vision_V18 (keepSynchronizedWithDisk=true) programFile=/programs/03 Sub Routines/Sub_Vision_V18.urp
  Folder PreSettings [hidden by the author, left out]
  '=========='
  Switch expression=Action
    Case (caseValue=13)
      SuppressedNode
        Folder Read [hidden by the author, left out]
    Case (caseValue=15)
      SuppressedNode
        Folder Detect [hidden by the author, left out]
    Case (caseValue=131)
      Folder Read (SensoPart)
        Action_Info := "search for landmark"
        CAM_LM := CAM_LMs[4]
        CAM_Relation := CAM_LM.capture_relation
        Folder go to capture pose [hidden by the author, left out]
        Loop While (checkContinuously=false) expression=not CAM_Done and  not ERROR.FLAG and  not CMD_Stop
          Folder adjust capture pose [hidden by the author, left out]
          Wait Sleep waitTime=2
          Folder trigger
            If ITM_ID≟1 and JIG≟7
              URCap VISOR Trigger (SensoPart VISOR Robotic, SensoPart Industriesensorik GmbH) dataModel(visorImageAcqSetup=2, visorId=0, visorSetJob=true, visorJobName=Landmark_INVITE_2); state(isChildrenLocked=true)
            ElseIf ITM_ID≟5 and JIG≟7
              URCap VISOR Trigger (SensoPart VISOR Robotic, SensoPart Industriesensorik GmbH) dataModel(visorImageAcqSetup=2, visorId=0, visorSetJob=true, visorJobName=Landmark_INVITE_2); state(isChildrenLocked=true)
            ElseIf ITM_ID≟13 and JIG≟7
              URCap VISOR Trigger (SensoPart VISOR Robotic, SensoPart Industriesensorik GmbH) dataModel(visorImageAcqSetup=2, visorId=0, visorSetJob=true, visorJobName=Landmark_INVITE_2); state(isChildrenLocked=true)
            ElseIf ITM_ID≟1 and JIG≟15
              URCap VISOR Trigger (SensoPart VISOR Robotic, SensoPart Industriesensorik GmbH) dataModel(visorImageAcqSetup=2, visorId=0, visorSetJob=true, visorJobName=QR_box); state(isChildrenLocked=true)
            ElseIf ITM_ID≟1 and JIG≟21
              URCap VISOR Trigger (SensoPart VISOR Robotic, SensoPart Industriesensorik GmbH) dataModel(visorImageAcqSetup=2, visorId=0, visorSetJob=true, visorJobName=PoTS); state(isChildrenLocked=true)
            ElseIf ITM_ID≟1 and JIG≟17
              URCap VISOR Trigger (SensoPart VISOR Robotic, SensoPart Industriesensorik GmbH) dataModel(visorImageAcqSetup=2, visorId=0, visorSetJob=true, visorJobName=Weigh_target); state(isChildrenLocked=true)
            SuppressedNode
              Folder init
                offset_result := visor_teachOffset(1,1,Base, 5000)
                Popup Message (haltProgram=false message=Supress This Folder inputType=Text)
            TM_3D_Found := visor_partsFound(1)
            If TM_3D_Found>0
              CAM_LM_Detected := True
              CAM_Captures := 0
            Else 
              CAM_LM_Detected := False
              CAM_Captures := CAM_Captures+1
            SuppressedNode
              CAM_LM_Deviatn := visor_getPose3d(1, 0)
            SuppressedNode
              If CAM_LM_Deviatn≠PSE_Z removedSiblings(If(type=Else checkContinuously=false, children(Assignment(valueSource=Expression, variable=CAM_LM_Detected, expression=False), Assignment(valueSource=Expression, variable=CAM_Captures, expression=CAM_Captures+1))))
                CAM_LM_Detected := True
                CAM_Captures := 0
          Folder result
            If CAM_LM_Detected
              If (CAM_LM_Refinmnt and CAM_LM_Refined) or  not CAM_LM_Refinmnt
                SuppressedNode
                  Switch expression=CAM_LM.id
                    Case (caseValue=1)
                      Folder Folder
                        'None'
                    Case (caseValue=2)
                      SuppressedNode
                        Folder SetUp
                          VEC_LM_PickUp := pose_trans(pose_inv(FRM_Reference), FRM_PickUp)
                      SuppressedNode
                        CAM_LM_Deviatn := pose_trans(pose_inv(FRM_PickUp), pose_trans(FRM_Reference, VEC_LM_PickUp))
                      SuppressedNode
                        FRM_PickUp := pose_trans(FRM_Reference, VEC_LM_PickUp)
                      SuppressedNode
                        Folder Frame test
                          PSE_T := p[0,0,0.03,d2r(-40),0,0]
                          PSE_A := p[0,0,0.15,d2r(-40),0,0]
                          MoveJ speed 60 deg/s, acceleration 80 deg/s^2 (useActiveTCP=false optimoveEnabled=false optiMoveSpeed=0.3 optiMoveAcceleration=0.09) tcp=TCP; feature=FRM_PickUp
                            Waypoint Variable (Variable): variable=PSE_A
                            Waypoint Variable (Variable): variable=PSE_T
                    Case (caseValue=3)
                      SuppressedNode
                        Folder SetUp
                          VEC_LM_DropOff1 := pose_trans(pose_inv(FRM_Reference), FRM_DropOff_1)
                      SuppressedNode
                        CAM_LM_Deviatn := pose_trans(pose_inv(FRM_DropOff_1), pose_trans(FRM_Reference, VEC_LM_DropOff1))
                      SuppressedNode
                        FRM_DropOff_1 := pose_trans(FRM_Reference, VEC_LM_DropOff1)
                      SuppressedNode
                        Folder Frame test
                          PSE_T := p[0,0,0.03,d2r(-40),0,0]
                          PSE_A := p[0,0,0.15,d2r(-40),0,0]
                          MoveJ speed 60 deg/s, acceleration 80 deg/s^2 (useActiveTCP=false optimoveEnabled=false optiMoveSpeed=0.3 optiMoveAcceleration=0.09) tcp=TCP; feature=FRM_DropOff_1
                            Waypoint Variable (Variable): variable=PSE_A
                            Waypoint Variable (Variable): variable=PSE_T
                    Case (caseValue=4)
                      SuppressedNode
                        Folder SetUp
                          VEC_LM_DropOff2 := pose_trans(pose_inv(FRM_Reference), FRM_DropOff_2)
                      SuppressedNode
                        CAM_LM_Deviatn := pose_trans(pose_inv(FRM_DropOff_2), pose_trans(FRM_Reference, VEC_LM_DropOff2))
                      SuppressedNode
                        FRM_DropOff_2 := pose_trans(FRM_Reference, VEC_LM_DropOff2)
                      SuppressedNode
                        Folder Frame test
                          PSE_T := p[0,0,0.03,0,0,0]
                          PSE_A := p[0,0,0.1,d2r(-45),0,0]
                          MoveJ speed 60 deg/s, acceleration 80 deg/s^2 (useActiveTCP=false optimoveEnabled=false optiMoveSpeed=0.3 optiMoveAcceleration=0.09) tcp=TCP; feature=FRM_DropOff_2
                            Waypoint Variable (Variable): variable=PSE_A
                            Waypoint Variable (Variable): variable=PSE_T
                    Case (caseValue=5)
                      SuppressedNode
                        Folder SetUp
                          VEC_LM_DropOff3 := pose_trans(pose_inv(FRM_Reference), FRM_DropOff_3)
                      SuppressedNode
                        FRM_DropOff_3 := pose_trans(FRM_Reference, VEC_LM_DropOff3)
                      SuppressedNode
                        Folder Frame test
                          PSE_T := p[0,0,0,0,0,0]
                          PSE_A := p[0,0,0.1,0,0,0]
                          MoveJ speed 60 deg/s, acceleration 80 deg/s^2 (useActiveTCP=false optimoveEnabled=false optiMoveSpeed=0.3 optiMoveAcceleration=0.09) tcp=TCP; feature=FRM_DropOff_3
                            Waypoint Variable (Variable): variable=PSE_A
                            Waypoint Variable (Variable): variable=PSE_T
                    Case (caseValue=6)
                      Folder Folder
                        'None'
                    Case (caseValue=7)
                      'Archive'
                    Case (caseValue=8)
                      SuppressedNode
                        Folder SetUp
                          VEC_LM_Centrifg := pose_trans(pose_inv(FRM_Reference), FRM_Centrifuge)
                      SuppressedNode
                        CAM_LM_Deviatn := pose_trans(pose_inv(FRM_Centrifuge), pose_trans(FRM_Reference, VEC_LM_Centrifg))
                      SuppressedNode
                        FRM_Centrifuge := pose_trans(FRM_Reference, VEC_LM_Centrifg)
                If ITM_ID≟1 and JIG≟7
                  CAM_LM_SSRack := visor_getPose3d(1, 0)
                ElseIf ITM_ID≟5 and JIG≟7
                  CAM_LM_SSRack := visor_getPose3d(1, 0)
                SuppressedNode
                  ElseIf ITM_ID≟13 and JIG≟7
                    CAM_LM_Bott := visor_getPose3d(1, 0)
                ElseIf ITM_ID≟1 and JIG≟15
                  CAM_LM_cont := visor_getPose3d(1, 0)
                  Trigger := get_actual_tcp_pose()
                ElseIf ITM_ID≟1 and JIG≟21
                  CAM_LM_cont := visor_getPose3d(1, 0)
                  Trigger := get_actual_tcp_pose()
                ElseIf ITM_ID≟1 and JIG≟17
                  CAM_LM_cont := visor_getPose3d(1, 0)
                  Trigger := get_actual_tcp_pose()
                CAM_Done := True
            ElseIf not CAM_LM_Detected and CAM_Captures<CAM_PRM_Retries
              CAM_LM_Refined := False
            ElseIf CAM_Captures≥CAM_PRM_Retries
              CAM_Done := True
              Folder Error
                Script: set_error(ERROR_NO_LANDMARK)
    Case (caseValue=151)
      Folder Detect (SensoPart) [hidden by the author, left out]
  '=========='
  Folder PostSettings [hidden by the author, left out]
SubProgram Sub_Action_V4 (keepSynchronizedWithDisk=false) programFile=/programs/03 Sub Routines/Sub_Action_V4.urp
  Folder PreSettings [hidden by the author, left out]
  '=========='
  Switch expression=Action
    Case (caseValue=1)
      Folder Pick
        Action_Info := "pick object"
        Script: do_transition(pose_trans(FRM_Reference, PSE_T), keep_rxry=OBJ_Picked)
        Folder EOAT
          If not OBJ_Picked
            Script: rq_move_and_wait_mm(GRP_Open_Pos)
        If PSE_A_H≠PSE_Z
          If JNT_Q≠JNT_Z
            Script: movej(get_inverse_kin(pose_trans(FRM_Reference, PSE_A_H), qnear=JNT_Q), r=0.050)
          Else 
            Script: movej(pose_trans(FRM_Reference, PSE_A_H), r=0.050)
        If PSE_A≠PSE_Z
          If JNT_Q≠JNT_Z
            Script: movej(get_inverse_kin(pose_trans(FRM_Reference, PSE_A), qnear=JNT_Q), r=0.020)
          Else 
            Script: movej(pose_trans(FRM_Reference, PSE_A), r=0.020)
        MoveL speed 400 mm/s, acceleration 500 mm/s^2 (useActiveTCP=true optimoveEnabled=false optiMoveSpeed=0.3 optiMoveAcceleration=0.09) feature=FRM_Reference
          If PSE_T_H≠PSE_Z
            Waypoint Variable (Variable): motionParameters(blendRadius=0.01); variable=PSE_T_H
          Waypoint Variable (Variable): motionParameters(jointSpeed=1.047198 jointAcceleration=1.396263 cartesianSpeed=0.12 cartesianAcceleration=0.08); variable=PSE_T
          Folder EOAT
            Script: rq_set_force_norm(50)
            Script: rq_close_and_wait()
            OBJ_Picked := rq_is_object_detected()
            If not OBJ_Picked
              Script: set_error(ERROR_NO_OBJECT_TO_PICK)
          Folder EXTT
            Switch expression=JIG
              Case (caseValue=1)
                Folder 3FG
                  If OBJ_Picked
                    Set DigitalOutput pin=GRP_3F_Open; digitalValue=1
          If PSE_R_H≠PSE_Z
            Waypoint Variable (Variable): motionParameters(blendRadius=0.01); variable=PSE_R
            Waypoint Variable (Variable): variable=PSE_R_H
          Else 
            Waypoint Variable (Variable): variable=PSE_R
    Case (caseValue=2)
      Folder Place [hidden by the author, left out]
    Case (caseValue=3)
      Folder Push
        Action_Info := "push"
    Case (caseValue=4)
      Folder Pull [hidden by the author, left out]
    SuppressedNode
      Case (caseValue=5)
        Placeholder
    Case (caseValue=6)
      Folder Drop the cap [hidden by the author, left out]
    Case (caseValue=7)
      Folder Load [hidden by the author, left out]
    Case (caseValue=8)
      Folder Unload [hidden by the author, left out]
    Case (caseValue=11)
      SuppressedNode
        Folder Place without opening gripper
          Action_Info := "place object without gripper opening"
          SuppressedNode
            Script: do_transition(pose_trans(FRM_Reference, PSE_T), keep_rxry=OBJ_Picked)
          Script: movel(FRM_Container_S, a=0.025, v=0.015, r=0.00001)
          Folder EXTT
            Switch expression=JIG
              Case (caseValue=1)
                Folder 3FG
                  If OBJ_Picked
                    Set DigitalOutput pin=GRP_3F_Open; digitalValue=1
          If PSE_A_H≠PSE_Z
            If JNT_Q≠JNT_Z
              Script: movej(get_inverse_kin(pose_trans(FRM_Reference, PSE_A_H), qnear=JNT_Q), r=0.050)
            Else 
              Script: movej(pose_trans(FRM_Reference, PSE_A_H), r=0.050)
          If PSE_A≠PSE_Z
            If JNT_Q≠JNT_Z
              Script: movej(get_inverse_kin(pose_trans(FRM_Reference, PSE_A), qnear=JNT_Q), r=0.020)
            Else 
              Script: movej(pose_trans(FRM_Reference, PSE_A), r=0.020)
          MoveL speed 400 mm/s, acceleration 500 mm/s^2 (useActiveTCP=true optimoveEnabled=false optiMoveSpeed=0.3 optiMoveAcceleration=0.09) feature=FRM_Reference
            If PSE_T_H≠PSE_Z
              Waypoint Variable (Variable): motionParameters(blendRadius=0.01); variable=PSE_T_H
            Waypoint Variable (Variable): motionParameters(jointSpeed=1.047198 jointAcceleration=1.396263 cartesianSpeed=0.09 cartesianAcceleration=0.05); variable=PSE_T
              Until TOOL_CONTACT_DETECTION (allowActions=false retraction=NONE decelerationAcceleration=0.5 decelerationAngularAcceleration=34.906585)
            Force Frame feature=FRM_Reference; selection=[1, 1, 1, 0, 0, 0]; wrench=[0, 0, 0, 0, 0, 0]; limitsForce=[0.1, 0.1, 0.01, 1.047198, 1.047198, 1.047198]; limitsMotion=[0.1, 0.1, 0.1, 0.349066, 0.349066, 0.349066]
              Waypoint Variable (Variable): motionParameters(jointSpeed=1.047198 jointAcceleration=1.396263 cartesianSpeed=0.07 cartesianAcceleration=0.04); variable=PSE_T
            Folder EXTT
              Switch expression=JIG
                Case (caseValue=1)
                  Folder 3FG
                    If OBJ_Picked
                      Set DigitalOutput pin=GRP_3F_Open; digitalValue=0
                      Wait Sleep waitTime=0.2
            Folder EOAT
              ''
    Case (caseValue=12)
      Folder Decap [hidden by the author, left out]
    Case (caseValue=13)
      Timer (action=Reset) variable(name=TMR_Barcode)
      Folder Read [hidden by the author, left out]
    Case (caseValue=15)
      Folder Detect
        Action_Info := "detect"
    Case (caseValue=30)
      Folder Shake [hidden by the author, left out]
    Case (caseValue=31)
      Action_Info := "Pick_Vial"
      Folder Pick_Vial [hidden by the author, left out]
    Case (caseValue=32)
      SuppressedNode
        decap := False
      Folder decap_Vial [hidden by the author, left out]
    Case (caseValue=33)
      Folder Shake and liquid transfer [hidden by the author, left out]
    SuppressedNode
      Case (caseValue=34)
        SafeHome (positionOptionType=SPEED_AND_ACCELERATION speed=1.047198 acceleration=1.396263 nextMotionTime=2)
        MoveJ speed 60 deg/s, acceleration 80 deg/s^2 (useActiveTCP=true optimoveEnabled=false optiMoveSpeed=0.3 optiMoveAcceleration=0.09) feature=Base
          Waypoint Waypoint_93: motionParameters(jointSpeed=0.436332 jointAcceleration=0.523599 cartesianSpeed=0.25 cartesianAcceleration=1.2); TCP in base x=206.301 y=-401.796 z=209.941 mm, rx=0 ry=0 rz=1.5608 rad; joints [-45.627, -84.145, -113.025, -72.821, 90.127, -225.014] deg; TCP offset x=0 y=0 z=161 mm, rx=3.1415 ry=0 rz=0 rad
        MoveL speed 250 mm/s, acceleration 1200 mm/s^2 (useActiveTCP=true optimoveEnabled=false optiMoveSpeed=0.3 optiMoveAcceleration=0.09) feature=Base
          Waypoint Waypoint_94: motionParameters(jointSpeed=1.047198 jointAcceleration=1.396263 cartesianSpeed=0.1 cartesianAcceleration=0.5); TCP in base x=200.866 y=-400.818 z=105.073 mm, rx=0 ry=0 rz=1.5608 rad; joints [-46.083, -90.669, -123.933, -55.389, 90.105, -225.416] deg
        URCap Gripper (Robotiq_Grippers, Robotiq Inc.) dataModel(position=100.0, force=27.84313725490196, speed=32.15686274509804, positionInDouble=100.0, forceInDouble=27.84313725490196, speedInDouble=32.15686274509804, slaveIds=[9], blocking=true)
        Wait Sleep waitTime=1
        MoveL speed 250 mm/s, acceleration 1200 mm/s^2 (useActiveTCP=true optimoveEnabled=false optiMoveSpeed=0.3 optiMoveAcceleration=0.09) feature=Base
          Waypoint Waypoint_95: motionParameters(jointSpeed=1.047198 jointAcceleration=1.396263 cartesianSpeed=0.1 cartesianAcceleration=0.5 blendRadius=0.05); TCP in base x=200.866 y=-400.818 z=325.177 mm, rx=0 ry=0 rz=1.5608 rad; joints [-46.018, -81.306, -98.396, -90.289, 90.129, -225.47] deg
        MoveJ speed 60 deg/s, acceleration 80 deg/s^2 (useActiveTCP=true optimoveEnabled=false optiMoveSpeed=0.3 optiMoveAcceleration=0.09) feature=Base
          Waypoint Waypoint_96: motionParameters(jointSpeed=0.436332 jointAcceleration=0.523599 cartesianSpeed=0.25 cartesianAcceleration=1.2 blendRadius=0.05); TCP in base x=-615.829 y=233.809 z=300 mm, rx=0.0051 ry=0.0087 rz=-2.1118 rad; joints [-188.832, -110.936, -69.076, -89.912, 89.674, -157.919] deg
        MoveL speed 250 mm/s, acceleration 1200 mm/s^2 (useActiveTCP=true optimoveEnabled=false optiMoveSpeed=0.3 optiMoveAcceleration=0.09) feature=Base
          Waypoint Waypoint_97: motionParameters(jointSpeed=1.047198 jointAcceleration=1.396263 cartesianSpeed=0.1 cartesianAcceleration=0.5); TCP in base x=-615.829 y=233.809 z=13.91 mm, rx=0.0051 ry=0.0087 rz=-2.1118 rad; joints [-188.874, -123.68, -94.539, -51.707, 89.657, -157.833] deg
        URCap Gripper (Robotiq_Grippers, Robotiq Inc.) dataModel(position=0.0, force=27.84313725490196, speed=32.15686274509804, positionInDouble=0.0, forceInDouble=27.84313725490196, speedInDouble=32.15686274509804, slaveIds=[9], blocking=true)
        MoveJ speed 60 deg/s, acceleration 80 deg/s^2 (useActiveTCP=true optimoveEnabled=false optiMoveSpeed=0.3 optiMoveAcceleration=0.09) feature=Base
          Waypoint Waypoint_98: motionParameters(jointSpeed=0.436332 jointAcceleration=0.523599 cartesianSpeed=0.25 cartesianAcceleration=1.2); TCP in base x=-615.829 y=233.809 z=300 mm, rx=0.0051 ry=0.0087 rz=-2.1118 rad; joints [-188.832, -110.936, -69.076, -89.912, 89.674, -157.919] deg
        SafeHome (positionOptionType=SPEED_AND_ACCELERATION speed=1.047198 acceleration=1.396263 nextMotionTime=2)
        SuppressedNode
          Folder Decap
            Action_Info := "decapping"
            Set DigitalOutput pin=GRP_3F_Enable; digitalValue=1
            Set DigitalOutput pin=GRP_3F_Decap; digitalValue=1
            Force Frame feature=Base; selection=[0, 0, 1, 0, 0, 0]; wrench=[0, 0, 1, 0, 0, 0]; limitsForce=[0.15, 0.15, 0.001, 1.047198, 1.047198, 1.047198]; limitsMotion=[0.1, 0.1, 0.1, 0.349066, 0.349066, 0.349066]
              Script: check_decapping(offset=0.015, timeout=10, abort=CMD_Hold)
            Set DigitalOutput pin=GRP_3F_Decap; digitalValue=0
            Set DigitalOutput pin=GRP_3F_Enable; digitalValue=0
            MoveL speed 250 mm/s, acceleration 1200 mm/s^2 (useActiveTCP=true optimoveEnabled=false optiMoveSpeed=0.3 optiMoveAcceleration=0.09) feature=Base
              Waypoint Waypoint_5: motionParameters(jointSpeed=1.047198 jointAcceleration=1.396263 cartesianSpeed=0.1 cartesianAcceleration=0.5 blendRadius=0.05); TCP in base x=-31.859 y=-349.402 z=312.809 mm, rx=0 ry=0 rz=0 rad; joints [-72.832, -66.838, -110.376, -92.778, 90.139, -162.834] deg
            MoveJ speed 60 deg/s, acceleration 80 deg/s^2 (useActiveTCP=true optimoveEnabled=false optiMoveSpeed=0.3 optiMoveAcceleration=0.09) feature=Base
              Waypoint cap_dump: motionParameters(jointSpeed=0.436332 jointAcceleration=0.523599 cartesianSpeed=0.25 cartesianAcceleration=1.2); TCP in base x=-139.169 y=-420.164 z=146.096 mm, rx=0 ry=0 rz=0 rad; joints [-90.79, -86.479, -121, -62.513, 90.12, -180.712] deg
            URCap Gripper (Robotiq_Grippers, Robotiq Inc.) dataModel(position=0.0, force=100.0, speed=100.0, positionInDouble=0.0, forceInDouble=100.0, speedInDouble=100.0, slaveIds=[9], blocking=true)
            MoveJ speed 60 deg/s, acceleration 80 deg/s^2 (useActiveTCP=true optimoveEnabled=false optiMoveSpeed=0.3 optiMoveAcceleration=0.09) feature=Base
              Waypoint Waypoint_5: motionParameters(jointSpeed=0.436332 jointAcceleration=0.523599 cartesianSpeed=0.25 cartesianAcceleration=1.2 blendRadius=0.05); TCP in base x=-31.859 y=-349.402 z=312.809 mm, rx=0 ry=0 rz=0 rad; joints [-72.832, -66.838, -110.376, -92.778, 90.139, -162.834] deg
            Set DigitalOutput pin=digital_out[5]; digitalValue=1
    SuppressedNode
      Case (caseValue=35)
        Folder Pick the powder container
          URCap VISOR Robotic App (SensoPart VISOR Robotic, SensoPart Industriesensorik GmbH) dataModel(visorAppTemplate=1); state(isChildrenLocked=true)
            URCap Easy Pick Setup (SensoPart VISOR Robotic, SensoPart Industriesensorik GmbH) dataModel(visorId=0, visorSetJob=true, visorJobName=Container_S, visorImageAcqSetup=2, visorCalibSetNo=7, visorDetector=1, visorImageAcqSource=1, visorOffsetSet=true, visorSetupStatus=3, Pose(key=visorImageAcqPose, Position(key=posePosition, Length(key=X value=-0.51041 unit=M), Length(key=Y value=0.417301 unit=M), Length(key=Z value=0.464095 unit=M)), Rotation(key=poseRotation, Angle(key=RX value=0.000026 unit=RAD), Angle(key=RY value=-0.000024 unit=RAD), Angle(key=RZ value=-2.896187 unit=RAD))), Pose(key=visorGripPose, Position(key=posePosition, Length(key=X value=-0.52891 unit=M), Length(key=Y value=0.461593 unit=M), Length(key=Z value=-0.178186 unit=M)), Rotation(key=poseRotation, Angle(key=RX value=-0.279814 unit=RAD), Angle(key=RY value=2.118244 unit=RAD), Angle(key=RZ value=-2.110314 unit=RAD)))); state(isChildrenLocked=true)
            URCap Process (SensoPart VISOR Robotic, SensoPart Industriesensorik GmbH) dataModel(Variable(key=visorCounterVar, variable(name=easyPickCount, initializeExpression=0)), Variable(key=visorPartsFoundVar, variable(name=easyPickParts, initializeExpression=0))); state(isChildrenLocked=true)
              URCap Image Acquisition Pose (SensoPart VISOR Robotic, SensoPart Industriesensorik GmbH) state(isChildrenLocked=true)
              URCap Object Detected (SensoPart VISOR Robotic, SensoPart Industriesensorik GmbH) state(isChildrenLocked=true)
                Folder Open Gripper
                  URCap Gripper (Robotiq_Grippers, Robotiq Inc.) dataModel(position=0.0, force=30.0, speed=40.0, positionInDouble=0.0, forceInDouble=30.0, speedInDouble=40.0, slaveIds=[9], blocking=true)
                  MoveJ speed 60 deg/s, acceleration 80 deg/s^2 (useActiveTCP=true optimoveEnabled=false optiMoveSpeed=0.3 optiMoveAcceleration=0.09) feature=Base
                    Waypoint Waypoint_13: TCP in base x=-479.451 y=284.141 z=125.27 mm, rx=-0.2768 ry=2.0984 rz=-2.1213 rad; joints [-165.671, -112.009, -127.874, -95.426, 1.192, -23.029] deg
                URCap Approach Pose (SensoPart VISOR Robotic, SensoPart Industriesensorik GmbH) dataModel(visorOffsetZ=-50.0); state(isChildrenLocked=true)
                URCap Target Pose (SensoPart VISOR Robotic, SensoPart Industriesensorik GmbH) state(isChildrenLocked=true)
                Folder Close Gripper
                  URCap Gripper (Robotiq_Grippers, Robotiq Inc.) dataModel(position=100.0, force=30.19607843137255, speed=40.0, positionInDouble=100.0, forceInDouble=30.19607843137255, speedInDouble=40.0, slaveIds=[9], blocking=true)
                URCap Exit Pose (SensoPart VISOR Robotic, SensoPart Industriesensorik GmbH) dataModel(visorOffsetZ=-50.0); state(isChildrenLocked=true)
              URCap No Object Detected (SensoPart VISOR Robotic, SensoPart Industriesensorik GmbH) dataModel(Variable(key=visorNoObjCountVar, variable(name=easyPickNoObj, initializeExpression=0)))
                Popup Message (haltProgram=false message=No Container detected inputType=Text)
          MoveJ speed 60 deg/s, acceleration 80 deg/s^2 (useActiveTCP=true optimoveEnabled=false optiMoveSpeed=0.3 optiMoveAcceleration=0.09) feature=Base
            SuppressedNode
              Waypoint Cont_midwa_1: motionParameters(jointSpeed=1.047198 jointAcceleration=1.396263 cartesianSpeed=0.25 cartesianAcceleration=1.2 blendRadius=0.01); TCP in base x=-462.252 y=294.856 z=204.322 mm, rx=-0.3472 ry=2.0343 rz=-2.0655 rad; joints [-166.773, -128.859, -129.893, 70.604, 5.32, -171.145] deg
            Waypoint Waypoint_70: motionParameters(jointSpeed=0.523599 jointAcceleration=0.698132 cartesianSpeed=0.25 cartesianAcceleration=1.2 blendRadius=0); TCP in base x=-472.821 y=292.44 z=207.418 mm, rx=-0.2598 ry=-2.0535 rz=2.0707 rad; joints [-170.164, -118.699, -96.461, -142.976, 25.725, -0.32] deg
            Waypoint Waypoint_78: motionParameters(jointSpeed=0.523599 jointAcceleration=0.872665 cartesianSpeed=0.25 cartesianAcceleration=1.2 blendRadius=0.05); TCP in base x=-51.45 y=-519.556 z=365.719 mm, rx=-1.2873 ry=1.0776 rz=-1.2185 rad; joints [-52.794, -108.287, -85.596, -162.721, 32.001, 1.948] deg
            Waypoint Waypoint_99: motionParameters(jointSpeed=0.523599 jointAcceleration=0.698132 cartesianSpeed=0.25 cartesianAcceleration=1.2 blendRadius=0.05); TCP in base x=-113.75 y=-390.11 z=317.307 mm, rx=-0.5194 ry=-0.8399 rz=1.7569 rad; joints [-108.345, -98.585, -86.606, -121.699, 124.957, 41.411] deg
          MoveL speed 250 mm/s, acceleration 1200 mm/s^2 (useActiveTCP=true optimoveEnabled=false optiMoveSpeed=0.3 optiMoveAcceleration=0.09) feature=Base
            Waypoint Waypoint_15: motionParameters(jointSpeed=1.047198 jointAcceleration=1.396263 cartesianSpeed=0.1 cartesianAcceleration=0.5 blendRadius=0.05); TCP in base x=29.144 y=-436.802 z=327.885 mm, rx=-0.5216 ry=-0.6236 rz=1.8627 rad; joints [-89.657, -89.204, -96.411, -97.086, 128.129, 64.023] deg
            Waypoint Waypoint_14: motionParameters(jointSpeed=1.047198 jointAcceleration=1.396263 cartesianSpeed=0.1 cartesianAcceleration=0.3); TCP in base x=68.712 y=-569.42 z=285.215 mm, rx=-0.6792 ry=-0.7121 rz=1.394 rad; joints [-90.137, -103.3, -96.148, -70.007, 141.633, 93.932] deg
            Waypoint Waypoint_100: motionParameters(jointSpeed=1.047198 jointAcceleration=1.396263 cartesianSpeed=0.05 cartesianAcceleration=0.3); TCP in base x=-47.22 y=-557.625 z=136.371 mm, rx=-0.6792 ry=-0.7121 rz=1.394 rad; joints [-101.643, -114.727, -100.71, -68.127, 140.302, 75.797] deg
          URCap Gripper (Robotiq_Grippers, Robotiq Inc.) dataModel(position=0.0, force=30.0, speed=40.0, positionInDouble=0.0, forceInDouble=30.0, speedInDouble=40.0, slaveIds=[9], blocking=true)
          MoveL speed 250 mm/s, acceleration 1200 mm/s^2 (useActiveTCP=true optimoveEnabled=false optiMoveSpeed=0.3 optiMoveAcceleration=0.09) feature=Base
            Waypoint Waypoint_25: motionParameters(jointSpeed=1.047198 jointAcceleration=1.396263 cartesianSpeed=0.1 cartesianAcceleration=0.3); TCP in base x=65.436 y=-569.388 z=287.821 mm, rx=-0.6792 ry=-0.7121 rz=1.394 rad; joints [-90.466, -103.248, -95.699, -70.925, 141.635, 93.398] deg
            Waypoint Waypoint_15: motionParameters(jointSpeed=1.047198 jointAcceleration=1.396263 cartesianSpeed=0.1 cartesianAcceleration=0.5 blendRadius=0.05); TCP in base x=29.144 y=-436.802 z=327.885 mm, rx=-0.5216 ry=-0.6236 rz=1.8627 rad; joints [-89.657, -89.204, -96.411, -97.086, 128.129, 64.023] deg
          SafeHome (positionOptionType=SPEED_AND_ACCELERATION speed=1.047198 acceleration=1.396263 nextMotionTime=2)
          SafeHome (positionOptionType=SPEED_AND_ACCELERATION speed=1.047198 acceleration=1.396263 nextMotionTime=2)
          SuppressedNode
            MoveJ speed 60 deg/s, acceleration 80 deg/s^2 (useActiveTCP=true optimoveEnabled=false optiMoveSpeed=0.3 optiMoveAcceleration=0.09) feature=Base
              Waypoint Container_midwa: motionParameters(blendRadius=0.05); TCP in base x=-379.239 y=-127.191 z=300 mm, rx=0 ry=0 rz=-1.2472 rad; joints [-141.945, -74.312, -107.466, -88.214, 90.137, -160.485] deg
          SuppressedNode
            URCap VISOR Robotic App (SensoPart VISOR Robotic, SensoPart Industriesensorik GmbH) dataModel(visorAppTemplate=1); state(isChildrenLocked=true)
              URCap Easy Pick Setup (SensoPart VISOR Robotic, SensoPart Industriesensorik GmbH) dataModel(visorId=0, visorSetJob=true, visorJobName=Target_container, visorImageAcqSetup=2, visorCalibSetNo=7, visorImageAcqSource=0, visorDetector=1, visorOffsetSet=true, visorSetupStatus=3, Pose(key=visorGripPose, Position(key=posePosition, Length(key=X value=-0.43018 unit=M), Length(key=Y value=0.500077 unit=M), Length(key=Z value=-0.155571 unit=M)), Rotation(key=poseRotation, Angle(key=RX value=0.000011 unit=RAD), Angle(key=RY value=0.000015 unit=RAD), Angle(key=RZ value=-2.896111 unit=RAD))), Pose(key=visorImageAcqPose, Position(key=posePosition, Length(key=X value=-0.391157 unit=M), Length(key=Y value=0.420635 unit=M), Length(key=Z value=0.411587 unit=M)), Rotation(key=poseRotation, Angle(key=RX value=-0.000006 unit=RAD), Angle(key=RY value=-0.000024 unit=RAD), Angle(key=RZ value=-2.896146 unit=RAD)))); state(isChildrenLocked=true)
              URCap Process (SensoPart VISOR Robotic, SensoPart Industriesensorik GmbH) dataModel(Variable(key=visorCounterVar, variable(name=easyPickCount_1, initializeExpression=0)), Variable(key=visorPartsFoundVar, variable(name=easyPickParts_1, initializeExpression=0))); state(isChildrenLocked=true)
                URCap Image Acquisition Pose (SensoPart VISOR Robotic, SensoPart Industriesensorik GmbH) state(isChildrenLocked=true)
                URCap Object Detected (SensoPart VISOR Robotic, SensoPart Industriesensorik GmbH) state(isChildrenLocked=true)
                  Folder Open Gripper
                    URCap Gripper (Robotiq_Grippers, Robotiq Inc.) dataModel(position=0.0, force=30.0, speed=40.0, positionInDouble=0.0, forceInDouble=30.0, speedInDouble=40.0, slaveIds=[9], blocking=true)
                  URCap Approach Pose (SensoPart VISOR Robotic, SensoPart Industriesensorik GmbH) dataModel(visorOffsetZ=-50.0); state(isChildrenLocked=true)
                  URCap Target Pose (SensoPart VISOR Robotic, SensoPart Industriesensorik GmbH) state(isChildrenLocked=true)
                  Folder Close Gripper
                    URCap Gripper (Robotiq_Grippers, Robotiq Inc.) dataModel(position=100.0, force=30.19607843137255, speed=40.0, positionInDouble=100.0, forceInDouble=30.19607843137255, speedInDouble=40.0, slaveIds=[9], blocking=true)
                  URCap Exit Pose (SensoPart VISOR Robotic, SensoPart Industriesensorik GmbH) dataModel(visorOffsetZ=-50.0); state(isChildrenLocked=true)
                URCap No Object Detected (SensoPart VISOR Robotic, SensoPart Industriesensorik GmbH) dataModel(Variable(key=visorNoObjCountVar, variable(name=easyPickNoObj_1, initializeExpression=0)))
                  Popup Message (haltProgram=false message=No Target container is detected inputType=Text)
          SuppressedNode
            MoveJ speed 60 deg/s, acceleration 80 deg/s^2 (useActiveTCP=true optimoveEnabled=false optiMoveSpeed=0.3 optiMoveAcceleration=0.09) feature=Base
              Waypoint Waypoint_16: motionParameters(jointSpeed=0.698132 jointAcceleration=0.872665 cartesianSpeed=0.25 cartesianAcceleration=1.2); TCP in base x=-389.004 y=141.378 z=266.753 mm, rx=0.0001 ry=-0.0001 rz=-2.8961 rad; joints [-181.152, -76.776, -110.541, -82.676, 90.144, -105.201] deg
              Waypoint Waypoint_17: motionParameters(jointSpeed=0.698132 jointAcceleration=0.872665 cartesianSpeed=0.25 cartesianAcceleration=1.2); TCP in base x=-35.034 y=-360.271 z=346.67 mm, rx=0.0001 ry=0 rz=-1.4195 rad; joints [-73.886, -68.929, -104.178, -96.885, 90.142, -82.58] deg
          SuppressedNode
            Set DigitalOutput pin=digital_out[5]; digitalValue=1
          SuppressedNode
            MoveL speed 250 mm/s, acceleration 1200 mm/s^2 (useActiveTCP=true optimoveEnabled=false optiMoveSpeed=0.3 optiMoveAcceleration=0.09) feature=Base
              Waypoint Waypoint_22: motionParameters(jointSpeed=1.047198 jointAcceleration=1.396263 cartesianSpeed=0.1 cartesianAcceleration=0.5); TCP in base x=-31.771 y=-348.512 z=220.918 mm, rx=0.0001 ry=0 rz=-1.1964 rad; joints [-72.82, -67.691, -123.366, -78.936, 90.15, -94.217] deg
              Waypoint Waypoint_23: motionParameters(jointSpeed=1.047198 jointAcceleration=1.396263 cartesianSpeed=0.05 cartesianAcceleration=0.3); TCP in base x=-31.891 y=-348.193 z=178.714 mm, rx=0.0001 ry=0 rz=-1.1964 rad; joints [-72.841, -69.405, -128.724, -71.864, 90.145, -94.213] deg
          SuppressedNode
            Set DigitalOutput pin=digital_out[5]; digitalValue=0
          SuppressedNode
            Wait Sleep waitTime=1
          SuppressedNode
            URCap Gripper (Robotiq_Grippers, Robotiq Inc.) dataModel(position=0.0, force=30.19607843137255, speed=40.0, positionInDouble=0.0, forceInDouble=30.19607843137255, speedInDouble=40.0, slaveIds=[9], blocking=true)
          SuppressedNode
            MoveL speed 250 mm/s, acceleration 1200 mm/s^2 (useActiveTCP=true optimoveEnabled=false optiMoveSpeed=0.3 optiMoveAcceleration=0.09) feature=Base
              Waypoint Waypoint_24: motionParameters(jointSpeed=1.047198 jointAcceleration=1.396263 cartesianSpeed=0.05 cartesianAcceleration=0.3); TCP in base x=-31.773 y=-348.52 z=270.997 mm, rx=0.0001 ry=0 rz=-1.1964 rad; joints [-72.799, -66.725, -116.549, -86.72, 90.151, -94.226] deg
          SuppressedNode
            SafeHome (positionOptionType=SPEED_AND_ACCELERATION speed=1.047198 acceleration=1.396263 nextMotionTime=2)
    SuppressedNode
      Case (caseValue=36)
        SuppressedNode
          MoveL speed 250 mm/s, acceleration 1200 mm/s^2 (useActiveTCP=true optimoveEnabled=false optiMoveSpeed=0.3 optiMoveAcceleration=0.09) feature=Base
            Waypoint Waypoint_26: TCP in base x=-30.182 y=-347.336 z=210.998 mm, rx=0 ry=0 rz=0 rad; joints [-72.486, -67.792, -124.787, -77.413, 90.141, -162.427] deg
        SuppressedNode
          URCap Gripper (Robotiq_Grippers, Robotiq Inc.) dataModel(position=100.0, force=30.19607843137255, speed=40.0, positionInDouble=100.0, forceInDouble=30.19607843137255, speedInDouble=40.0, slaveIds=[9], blocking=true)
        SuppressedNode
          Folder Decap
            Action_Info := "decapping"
            Set DigitalOutput pin=GRP_3F_Enable; digitalValue=1
            Set DigitalOutput pin=GRP_3F_Decap; digitalValue=1
            Force Frame feature=Base; selection=[0, 0, 1, 0, 0, 0]; wrench=[0, 0, 1, 0, 0, 0]; limitsForce=[0.15, 0.15, 0.001, 1.047198, 1.047198, 1.047198]; limitsMotion=[0.1, 0.1, 0.1, 0.349066, 0.349066, 0.349066]
              Script: check_decapping(offset=0.015, timeout=12, abort=CMD_Hold)
            Set DigitalOutput pin=GRP_3F_Decap; digitalValue=0
            Set DigitalOutput pin=GRP_3F_Enable; digitalValue=0
            MoveL speed 250 mm/s, acceleration 1200 mm/s^2 (useActiveTCP=true optimoveEnabled=false optiMoveSpeed=0.3 optiMoveAcceleration=0.09) feature=Base
              Waypoint Waypoint_27: motionParameters(jointSpeed=1.047198 jointAcceleration=1.396263 cartesianSpeed=0.1 cartesianAcceleration=0.5 blendRadius=0.05); TCP in base x=-30.361 y=-347.415 z=279.539 mm, rx=0 ry=0 rz=-0.0004 rad; joints [-72.488, -66.465, -115.449, -88.079, 90.139, -162.449] deg
              Waypoint Waypoint_28: motionParameters(jointSpeed=1.047198 jointAcceleration=1.396263 cartesianSpeed=0.1 cartesianAcceleration=0.5 blendRadius=0.05); TCP in base x=-154.725 y=-473.257 z=246.189 mm, rx=0 ry=0 rz=-0.0004 rad; joints [-92.526, -89.454, -102.579, -77.959, 90.132, -182.495] deg
              Waypoint Waypoint_29: motionParameters(jointSpeed=1.047198 jointAcceleration=1.396263 cartesianSpeed=0.1 cartesianAcceleration=0.3); TCP in base x=-145.695 y=-485.909 z=46.677 mm, rx=0 ry=0 rz=-0.0004 rad; joints [-91.444, -104.036, -119.144, -46.812, 90.094, -181.324] deg
            URCap Gripper (Robotiq_Grippers, Robotiq Inc.) dataModel(position=61.24306326304106, force=30.19607843137255, speed=40.0, positionInDouble=61.24306326304106, forceInDouble=30.19607843137255, speedInDouble=40.0, slaveIds=[9], blocking=true)
            MoveL speed 250 mm/s, acceleration 1200 mm/s^2 (useActiveTCP=true optimoveEnabled=false optiMoveSpeed=0.3 optiMoveAcceleration=0.09) feature=Base
              Waypoint Waypoint_38: motionParameters(jointSpeed=1.047198 jointAcceleration=1.396263 cartesianSpeed=0.1 cartesianAcceleration=0.5 blendRadius=0.05); TCP in base x=-145.695 y=-485.909 z=261.43 mm, rx=0 ry=0 rz=-0.0004 rad; joints [-91.4, -90.37, -99.399, -80.223, 90.132, -181.38] deg
              URCap Gripper (Robotiq_Grippers, Robotiq Inc.) dataModel(position=0.0, force=30.19607843137255, speed=40.0, positionInDouble=0.0, forceInDouble=30.19607843137255, speedInDouble=40.0, slaveIds=[9], blocking=true)
              Waypoint Waypoint_30: motionParameters(jointSpeed=1.047198 jointAcceleration=1.396263 cartesianSpeed=0.1 cartesianAcceleration=0.5 blendRadius=0.05); TCP in base x=-30.182 y=-347.336 z=265.578 mm, rx=0 ry=0 rz=0 rad; joints [-72.462, -66.558, -117.437, -85.997, 90.142, -162.436] deg
              Waypoint Waypoint_31: motionParameters(jointSpeed=1.047198 jointAcceleration=1.396263 cartesianSpeed=0.1 cartesianAcceleration=0.5); TCP in base x=-30.182 y=-347.336 z=175.833 mm, rx=0 ry=0 rz=0 rad; joints [-72.5, -69.38, -129.182, -71.43, 90.136, -162.42] deg
            URCap Gripper (Robotiq_Grippers, Robotiq Inc.) dataModel(position=79.44506104328524, force=30.19607843137255, speed=40.0, positionInDouble=79.44506104328524, forceInDouble=30.19607843137255, speedInDouble=40.0, slaveIds=[9], blocking=true)
            Wait Sleep waitTime=1
            Set DigitalOutput pin=digital_out[5]; digitalValue=1
            MoveL speed 250 mm/s, acceleration 1200 mm/s^2 (useActiveTCP=true optimoveEnabled=false optiMoveSpeed=0.3 optiMoveAcceleration=0.09) feature=Base
              Waypoint Waypoint_32: motionParameters(jointSpeed=1.047198 jointAcceleration=1.396263 cartesianSpeed=0.1 cartesianAcceleration=0.5 blendRadius=0.05); TCP in base x=-30.182 y=-347.336 z=316.067 mm, rx=0 ry=0 rz=0 rad; joints [-72.438, -66.521, -110.081, -93.39, 90.138, -162.442] deg
            URCap VISOR Robotic App (SensoPart VISOR Robotic, SensoPart Industriesensorik GmbH) dataModel(visorAppTemplate=1); state(isChildrenLocked=true)
              URCap Easy Pick Setup (SensoPart VISOR Robotic, SensoPart Industriesensorik GmbH) dataModel(visorId=0, visorSetJob=true, visorJobName=Weigh_scale, visorImageAcqSetup=2, visorImageAcqSource=1, visorCalibSetNo=9, visorDetector=1, visorSetupStatus=5, visorOffsetSet=true, Pose(key=visorGripPose, Position(key=posePosition, Length(key=X value=-0.66092 unit=M), Length(key=Y value=-0.026261 unit=M), Length(key=Z value=0.113423 unit=M)), Rotation(key=poseRotation, Angle(key=RX value=0.044036 unit=RAD), Angle(key=RY value=-0.006733 unit=RAD), Angle(key=RZ value=-1.658906 unit=RAD)))); state(isChildrenLocked=true)
              URCap Process (SensoPart VISOR Robotic, SensoPart Industriesensorik GmbH) dataModel(Variable(key=visorCounterVar, variable(name=easyPickCount_2, initializeExpression=0)), Variable(key=visorPartsFoundVar, variable(name=easyPickParts_2, initializeExpression=0))); state(isChildrenLocked=true)
                URCap Image Acquisition Pose (SensoPart VISOR Robotic, SensoPart Industriesensorik GmbH) state(isChildrenLocked=true)
                URCap Object Detected (SensoPart VISOR Robotic, SensoPart Industriesensorik GmbH) state(isChildrenLocked=true)
                  Folder Open Gripper
                    Wait NoWait
                  URCap Approach Pose (SensoPart VISOR Robotic, SensoPart Industriesensorik GmbH) dataModel(visorOffsetZ=-50.0); state(isChildrenLocked=true)
                  URCap Target Pose (SensoPart VISOR Robotic, SensoPart Industriesensorik GmbH) state(isChildrenLocked=true)
                  Folder Close Gripper
                    URCap Gripper (Robotiq_Grippers, Robotiq Inc.) dataModel(position=0.0, force=30.19607843137255, speed=40.0, positionInDouble=0.0, forceInDouble=30.19607843137255, speedInDouble=40.0, slaveIds=[9], blocking=true)
                  URCap Exit Pose (SensoPart VISOR Robotic, SensoPart Industriesensorik GmbH) dataModel(visorOffsetZ=-100.0); state(isChildrenLocked=true)
                URCap No Object Detected (SensoPart VISOR Robotic, SensoPart Industriesensorik GmbH) dataModel(Variable(key=visorNoObjCountVar, variable(name=easyPickNoObj_2, initializeExpression=0)))
                  Popup Message (haltProgram=false message=No weigh scale is detected inputType=Text)
            SafeHome (positionOptionType=SPEED_AND_ACCELERATION speed=1.047198 acceleration=1.396263 nextMotionTime=2)
            MoveJ speed 60 deg/s, acceleration 80 deg/s^2 (useActiveTCP=true optimoveEnabled=false optiMoveSpeed=0.3 optiMoveAcceleration=0.09) feature=Base
              Waypoint Waypoint_39: TCP in base x=137.772 y=-577.76 z=300 mm, rx=0 ry=0 rz=-1.5944 rad; joints [-63.54, -101.785, -81.001, -87.198, 90.144, -62.245] deg
            MoveL speed 250 mm/s, acceleration 1200 mm/s^2 (useActiveTCP=true optimoveEnabled=false optiMoveSpeed=0.3 optiMoveAcceleration=0.09) feature=Base
              Waypoint Waypoint_41: motionParameters(jointSpeed=1.047198 jointAcceleration=1.396263 cartesianSpeed=0.1 cartesianAcceleration=0.5); TCP in base x=74.223 y=-565.642 z=234.62 mm, rx=-0.5169 ry=0.5292 rz=-1.5296 rad; joints [-54.985, -107.527, -85.329, -102.066, 60.279, -46.981] deg
              Waypoint Waypoint_40: motionParameters(jointSpeed=1.047198 jointAcceleration=1.396263 cartesianSpeed=0.05 cartesianAcceleration=0.3); TCP in base x=39.988 y=-564.833 z=191.055 mm, rx=-0.7676 ry=0.3431 rz=-2.2413 rad; joints [-57.701, -107.406, -92.471, -93.607, 59.17, -6.639] deg
            URCap Gripper (Robotiq_Grippers, Robotiq Inc.) dataModel(position=100.0, force=20.0, speed=30.0, positionInDouble=100.0, forceInDouble=20.0, speedInDouble=30.0, slaveIds=[9], blocking=true)
            Loop Counting (count=2) loopVariable(name=Loop_2)
              MoveL speed 250 mm/s, acceleration 1200 mm/s^2 (useActiveTCP=true optimoveEnabled=false optiMoveSpeed=0.3 optiMoveAcceleration=0.09) feature=Base
                Waypoint Waypoint_42: motionParameters(jointSpeed=1.047198 jointAcceleration=1.396263 cartesianSpeed=0.5 cartesianAcceleration=1.2 blendRadius=0); TCP in base x=41.363 y=-564.865 z=192.806 mm, rx=0.2785 ry=0.6241 rz=0.7623 rad; joints [-57.586, -107.397, -92.198, -93.963, 59.209, -186.442] deg
                Waypoint Waypoint_43: TCP in base x=41.363 y=-564.865 z=192.806 mm, rx=0.9734 ry=0.0641 rz=2.8083 rad; joints [-57.585, -107.391, -92.207, -93.949, 59.207, -310.817] deg
              URCap Gripper (Robotiq_Grippers, Robotiq Inc.) dataModel(position=24.83906770255271, force=20.0, speed=30.19607843137255, positionInDouble=24.83906770255271, forceInDouble=20.0, speedInDouble=30.19607843137255, slaveIds=[9], blocking=true)
              MoveL speed 250 mm/s, acceleration 1200 mm/s^2 (useActiveTCP=true optimoveEnabled=false optiMoveSpeed=0.3 optiMoveAcceleration=0.09) feature=Base
                Waypoint Waypoint_44: motionParameters(jointSpeed=1.047198 jointAcceleration=1.396263 cartesianSpeed=0.5 cartesianAcceleration=1.2 blendRadius=0); TCP in base x=40.883 y=-564.854 z=192.194 mm, rx=0.1109 ry=0.6592 rz=0.2757 rad; joints [-57.626, -107.402, -92.291, -93.842, 59.196, -157.494] deg
                Waypoint Waypoint_45: TCP in base x=42.648 y=-564.896 z=194.439 mm, rx=-0.4517 ry=0.5632 rz=-1.3434 rad; joints [-57.484, -107.381, -91.951, -94.273, 59.256, -60.779] deg
              URCap Gripper (Robotiq_Grippers, Robotiq Inc.) dataModel(position=78.43137254901961, force=20.0, speed=30.0, positionInDouble=78.43137254901961, forceInDouble=20.0, speedInDouble=30.0, slaveIds=[9], blocking=true)
            MoveL speed 250 mm/s, acceleration 1200 mm/s^2 (useActiveTCP=true optimoveEnabled=false optiMoveSpeed=0.3 optiMoveAcceleration=0.09) feature=Base
              Waypoint Waypoint_46: motionParameters(jointSpeed=1.047198 jointAcceleration=1.396263 cartesianSpeed=0.05 cartesianAcceleration=0.3); TCP in base x=99.944 y=-566.244 z=267.343 mm, rx=-0.4517 ry=0.5632 rz=-1.3434 rad; joints [-53.041, -108.287, -79.23, -108.385, 61.102, -56.184] deg
              Waypoint Waypoint_47: motionParameters(jointSpeed=1.047198 jointAcceleration=1.396263 cartesianSpeed=0.1 cartesianAcceleration=0.5 blendRadius=0); TCP in base x=99.944 y=-566.244 z=267.343 mm, rx=-0.1017 ry=0.0587 rz=-1.4579 rad; joints [-63.671, -99.121, -88.981, -82.751, 84.056, -70.038] deg
              Waypoint Waypoint_48: motionParameters(jointSpeed=1.047198 jointAcceleration=1.396263 cartesianSpeed=0.25 cartesianAcceleration=1.2); TCP in base x=-136.183 y=-647.487 z=294.248 mm, rx=-0.1017 ry=0.0587 rz=-1.4579 rad; joints [-87.788, -109.526, -72.49, -86.263, 84.243, -94.331] deg
              Waypoint Waypoint_49: TCP in base x=-159.024 y=-641.021 z=47.692 mm, rx=0 ry=0 rz=-1.4579 rad; joints [-92.238, -121.266, -92.571, -56.15, 90.14, -98.675] deg
            URCap Gripper (Robotiq_Grippers, Robotiq Inc.) dataModel(position=33.9400665926748, force=20.0, speed=30.19607843137255, positionInDouble=33.9400665926748, forceInDouble=20.0, speedInDouble=30.19607843137255, slaveIds=[9], blocking=true)
            MoveL speed 250 mm/s, acceleration 1200 mm/s^2 (useActiveTCP=true optimoveEnabled=false optiMoveSpeed=0.3 optiMoveAcceleration=0.09) feature=Base
              Waypoint Waypoint_50: TCP in base x=-159.024 y=-641.021 z=291.114 mm, rx=0 ry=0 rz=-1.4579 rad; joints [-92.2, -111.308, -69.838, -88.841, 90.151, -98.75] deg
              SafeHome (positionOptionType=SPEED_AND_ACCELERATION speed=1.047198 acceleration=1.396263 nextMotionTime=2)
    SuppressedNode
      Case (caseValue=37)
        SuppressedNode
          URCap VISOR Robotic App (SensoPart VISOR Robotic, SensoPart Industriesensorik GmbH) dataModel(visorAppTemplate=1); state(isChildrenLocked=true)
            URCap Easy Pick Setup (SensoPart VISOR Robotic, SensoPart Industriesensorik GmbH) dataModel(visorId=0, visorSetJob=true, visorJobName=Spatula, visorImageAcqSetup=2, visorImageAcqSource=1, visorCalibSetNo=10, visorDetector=1, visorOffsetSet=true, visorSetupStatus=5, Pose(key=visorGripPose, Position(key=posePosition, Length(key=X value=-0.64401 unit=M), Length(key=Y value=-0.309906 unit=M), Length(key=Z value=0.133972 unit=M)), Rotation(key=poseRotation, Angle(key=RX value=0.000082 unit=RAD), Angle(key=RY value=0.000005 unit=RAD), Angle(key=RZ value=3.001273 unit=RAD)))); state(isChildrenLocked=true)
            URCap Process (SensoPart VISOR Robotic, SensoPart Industriesensorik GmbH) dataModel(Variable(key=visorCounterVar, variable(name=easyPickCount_3, initializeExpression=0)), Variable(key=visorPartsFoundVar, variable(name=easyPickParts_3, initializeExpression=0))); state(isChildrenLocked=true)
              URCap Image Acquisition Pose (SensoPart VISOR Robotic, SensoPart Industriesensorik GmbH) state(isChildrenLocked=true)
              URCap Object Detected (SensoPart VISOR Robotic, SensoPart Industriesensorik GmbH) state(isChildrenLocked=true)
                Folder Open Gripper
                  URCap Gripper (Robotiq_Grippers, Robotiq Inc.) dataModel(position=0.0, force=20.0, speed=30.19607843137255, positionInDouble=0.0, forceInDouble=20.0, speedInDouble=30.19607843137255, slaveIds=[9], blocking=true)
                URCap Approach Pose (SensoPart VISOR Robotic, SensoPart Industriesensorik GmbH) dataModel(visorOffsetZ=-100.0); state(isChildrenLocked=true)
                URCap Target Pose (SensoPart VISOR Robotic, SensoPart Industriesensorik GmbH) state(isChildrenLocked=true)
                Folder Close Gripper
                  URCap Gripper (Robotiq_Grippers, Robotiq Inc.) dataModel(position=100.0, force=20.0, speed=30.19607843137255, positionInDouble=100.0, forceInDouble=20.0, speedInDouble=30.19607843137255, slaveIds=[9], blocking=true)
                URCap Exit Pose (SensoPart VISOR Robotic, SensoPart Industriesensorik GmbH) dataModel(visorToolSpeed=100.0, visorToolAcc=300.0, visorOffsetZ=-200.0); state(isChildrenLocked=true)
              URCap No Object Detected (SensoPart VISOR Robotic, SensoPart Industriesensorik GmbH) dataModel(Variable(key=visorNoObjCountVar, variable(name=easyPickNoObj_3, initializeExpression=0)))
                Popup Message (haltProgram=false message=No spatula is detected inputType=Text)
        URCap VISOR Robotic App (SensoPart VISOR Robotic, SensoPart Industriesensorik GmbH) dataModel(visorAppTemplate=1); state(isChildrenLocked=true)
          URCap Easy Pick Setup (SensoPart VISOR Robotic, SensoPart Industriesensorik GmbH) dataModel(visorId=0, visorSetJob=true, visorJobName=Spatula_horizontal, visorImageAcqSetup=2, visorImageAcqSource=0, visorDetector=1, visorOffsetSet=true, visorSetupStatus=1, Pose(key=visorImageAcqPose, Position(key=posePosition, Length(key=X value=-0.477866 unit=M), Length(key=Y value=0.377208 unit=M), Length(key=Z value=0.48314 unit=M)), Rotation(key=poseRotation, Angle(key=RX value=-0.000072 unit=RAD), Angle(key=RY value=-0.000033 unit=RAD), Angle(key=RZ value=-1.610249 unit=RAD))), Pose(key=visorGripPose, Position(key=posePosition, Length(key=X value=-0.547139 unit=M), Length(key=Y value=0.33515 unit=M), Length(key=Z value=0.041533 unit=M)), Rotation(key=poseRotation, Angle(key=RX value=2.188123 unit=RAD), Angle(key=RY value=-0.020843 unit=RAD), Angle(key=RZ value=2.219811 unit=RAD)))); state(isChildrenLocked=true)
          URCap Process (SensoPart VISOR Robotic, SensoPart Industriesensorik GmbH) dataModel(Variable(key=visorCounterVar, variable(name=easyPickCount_5, initializeExpression=0)), Variable(key=visorPartsFoundVar, variable(name=easyPickParts_5, initializeExpression=0))); state(isChildrenLocked=true)
            URCap Image Acquisition Pose (SensoPart VISOR Robotic, SensoPart Industriesensorik GmbH) state(isChildrenLocked=true)
            URCap Object Detected (SensoPart VISOR Robotic, SensoPart Industriesensorik GmbH) state(isChildrenLocked=true)
              Folder Open Gripper
                URCap Gripper (Robotiq_Grippers, Robotiq Inc.) dataModel(position=43.04106548279689, force=30.0, speed=30.0, positionInDouble=43.04106548279689, forceInDouble=30.0, speedInDouble=30.0, slaveIds=[9], blocking=true)
              URCap Approach Pose (SensoPart VISOR Robotic, SensoPart Industriesensorik GmbH) dataModel(visorOffsetZ=-130.0); state(isChildrenLocked=true)
              URCap Target Pose (SensoPart VISOR Robotic, SensoPart Industriesensorik GmbH) state(isChildrenLocked=true)
              Folder Close Gripper
                URCap Gripper (Robotiq_Grippers, Robotiq Inc.) dataModel(position=100.0, force=30.0, speed=30.0, positionInDouble=100.0, forceInDouble=30.0, speedInDouble=30.0, slaveIds=[9], blocking=true)
              URCap Exit Pose (SensoPart VISOR Robotic, SensoPart Industriesensorik GmbH) dataModel(visorOffsetZ=-170.0); state(isChildrenLocked=true)
            URCap No Object Detected (SensoPart VISOR Robotic, SensoPart Industriesensorik GmbH) dataModel(Variable(key=visorNoObjCountVar, variable(name=easyPickNoObj_5, initializeExpression=0)))
              Popup Message (haltProgram=false message=No Spatula detected inputType=Text)
        SuppressedNode
          MoveJ speed 60 deg/s, acceleration 80 deg/s^2 (useActiveTCP=true optimoveEnabled=false optiMoveSpeed=0.3 optiMoveAcceleration=0.09) feature=Base
            Waypoint Waypoint_1: motionParameters(jointSpeed=1.047198 jointAcceleration=1.396263 cartesianSpeed=0.1 cartesianAcceleration=0.5 blendRadius=0.05); TCP in base x=-359.544 y=319.273 z=259.271 mm, rx=2.1553 ry=-0.0199 rz=2.2443 rad; joints [-228.189, -86.975, -126.838, -149.463, 223.669, -271.634] deg
            Waypoint Waypoint_51: motionParameters(jointSpeed=1.047198 jointAcceleration=1.396263 cartesianSpeed=0.1 cartesianAcceleration=0.5 blendRadius=0); TCP in base x=-477.866 y=377.208 z=483.14 mm, rx=-0.0001 ry=0 rz=-1.6102 rad; joints [-205.499, -110.086, -42.439, -117.467, 90.106, -203.428] deg
            Waypoint Waypoint_52: TCP in base x=-42.31 y=-356.333 z=399.894 mm, rx=0 ry=0 rz=-0.1228 rad; joints [-74.871, -69.823, -95.716, -104.453, 90.124, -157.892] deg
        MoveL speed 50 mm/s, acceleration 300 mm/s^2 (useActiveTCP=true optimoveEnabled=false optiMoveSpeed=0.3 optiMoveAcceleration=0.09) feature=Base
          Waypoint Waypoint_3: motionParameters(jointSpeed=1.047198 jointAcceleration=1.396263 cartesianSpeed=0.05 cartesianAcceleration=0.3); TCP in base x=-31.864 y=-349.975 z=230.259 mm, rx=0 ry=0 rz=0 rad; joints [-72.901, -67.669, -121.993, -80.33, 90.142, -162.853] deg
          Waypoint Waypoint_80: motionParameters(jointSpeed=1.047198 jointAcceleration=1.396263 cartesianSpeed=0.05 cartesianAcceleration=0.3); TCP in base x=143.03 y=-569.853 z=275.754 mm, rx=1.2979 ry=0.0264 rz=2.7129 rad; joints [-47.784, -117.454, -67.716, -126.008, 56.917, 63.329] deg
          Loop Counting (count=3) loopVariable(name=Loop_3)
            Waypoint Waypoint_55: motionParameters(jointSpeed=1.047198 jointAcceleration=1.396263 cartesianSpeed=0.05 cartesianAcceleration=0.3); TCP in base x=73.857 y=-577.013 z=221.505 mm, rx=1.2979 ry=0.0264 rz=2.7129 rad; joints [-52.913, -114.774, -80.289, -113.397, 53.656, 58.584] deg
              Until TOOL_CONTACT_DETECTION (allowActions=false retraction=0 decelerationAcceleration=3 decelerationAngularAcceleration=34.906585)
            Waypoint Waypoint_56: motionParameters(jointSpeed=1.047198 jointAcceleration=1.396263 cartesianSpeed=0.05 cartesianAcceleration=0.3); TCP in base x=135.677 y=-579.448 z=242.231 mm, rx=1.5554 ry=0.0154 rz=2.5559 rad; joints [-47.427, -124.812, -65.265, -134.284, 52.841, 72.036] deg
          Loop Counting (count=2) loopVariable(name=Loop_5)
            Waypoint Waypoint_56: motionParameters(jointSpeed=1.047198 jointAcceleration=1.396263 cartesianSpeed=0.05 cartesianAcceleration=0.3); TCP in base x=135.677 y=-579.448 z=242.231 mm, rx=1.5554 ry=0.0154 rz=2.5559 rad; joints [-47.427, -124.812, -65.265, -134.284, 52.841, 72.036] deg
            Waypoint Waypoint_101: motionParameters(jointSpeed=1.047198 jointAcceleration=1.396263 cartesianSpeed=0.5 cartesianAcceleration=1.2); TCP in base x=143.391 y=-581.809 z=226.065 mm, rx=1.6397 ry=0.0079 rz=2.5024 rad; joints [-46.773, -128.399, -63.349, -137.511, 52.317, 75.293] deg
          Waypoint Waypoint_59: motionParameters(jointSpeed=1.047198 jointAcceleration=1.396263 cartesianSpeed=0.05 cartesianAcceleration=0.3); TCP in base x=272.401 y=-578.183 z=239.561 mm, rx=2.127 ry=0.1139 rz=2.1556 rad; joints [-37.816, -154.733, -25.502, -178.522, 53.445, 96.624] deg
          Waypoint Waypoint_58: motionParameters(jointSpeed=1.047198 jointAcceleration=1.396263 cartesianSpeed=0.05 cartesianAcceleration=0.3); TCP in base x=223.649 y=-578.478 z=276.546 mm, rx=2.1743 ry=-0.0441 rz=2.0587 rad; joints [-41.771, -153.265, -25.455, -184.54, 55.381, 96.631] deg
        MoveJ speed 30 deg/s, acceleration 50 deg/s^2 (useActiveTCP=true optimoveEnabled=false optiMoveSpeed=0.3 optiMoveAcceleration=0.09) feature=Base
          Waypoint Waypoint_60: motionParameters(jointSpeed=0.349066 jointAcceleration=0.523599 cartesianSpeed=0.25 cartesianAcceleration=1.2 blendRadius=0.05); TCP in base x=-13.316 y=-544.772 z=383.372 mm, rx=2.2082 ry=0.0375 rz=2.0976 rad; joints [-53.447, -120.321, -68.514, -175.377, 39.556, 98.101] deg
          Waypoint Waypoint_61: motionParameters(jointSpeed=0.349066 jointAcceleration=0.523599 cartesianSpeed=0.25 cartesianAcceleration=1.2 blendRadius=0.05); TCP in base x=-412.189 y=-356.447 z=383.372 mm, rx=1.7517 ry=-0.74 rz=1.6007 rad; joints [-101.195, -120.321, -68.514, -175.377, 39.556, 98.101] deg
          Waypoint Waypoint_62: motionParameters(jointSpeed=0.349066 jointAcceleration=0.523599 cartesianSpeed=0.25 cartesianAcceleration=1.2); TCP in base x=-542.659 y=-114.282 z=251.262 mm, rx=1.813 ry=-0.6794 rz=1.6553 rad; joints [-123.661, -111.262, -103.952, -159.22, 12.548, 108.767] deg
        MoveL speed 250 mm/s, acceleration 1200 mm/s^2 (useActiveTCP=true optimoveEnabled=false optiMoveSpeed=0.3 optiMoveAcceleration=0.09) feature=Base
          Waypoint Waypoint_63: motionParameters(jointSpeed=1.047198 jointAcceleration=1.396263 cartesianSpeed=0.05 cartesianAcceleration=0.3); TCP in base x=-532.496 y=-127.81 z=159.342 mm, rx=1.813 ry=-0.6794 rz=1.6553 rad; joints [-121.654, -119.526, -108.357, -144.665, 14.532, 106.823] deg
          Waypoint Waypoint_102: motionParameters(jointSpeed=1.047198 jointAcceleration=1.396263 cartesianSpeed=0.05 cartesianAcceleration=0.3); TCP in base x=-576.035 y=-66.27 z=306.74 mm, rx=0.8621 ry=-0.2554 rz=2.1952 rad; joints [-142.141, -87.685, -107.535, -64.498, 50.077, -8.596] deg
          Waypoint Waypoint_103: motionParameters(jointSpeed=1.047198 jointAcceleration=1.396263 cartesianSpeed=0.05 cartesianAcceleration=0.3); TCP in base x=-581.965 y=-59.291 z=312.082 mm, rx=0.8621 ry=-0.2554 rz=2.1952 rad; joints [-143.275, -88.018, -106.65, -64.116, 50.29, -10.05] deg
          Waypoint Waypoint_81: motionParameters(jointSpeed=1.047198 jointAcceleration=1.396263 cartesianSpeed=0.5 cartesianAcceleration=1.2); TCP in base x=-581.965 y=-59.291 z=290.576 mm, rx=0.8621 ry=-0.2554 rz=2.1952 rad; joints [-143.281, -88.87, -109.094, -60.824, 50.286, -10.043] deg
          Waypoint Decap_above: TCP in base x=-31.864 y=-349.975 z=288.042 mm, rx=0 ry=0 rz=0 rad; joints [-72.875, -66.865, -113.978, -89.149, 90.141, -162.862] deg
